DATA_BLOCK "DI_GC02_FB06_Conv_G115D"
{ S7_Optimized_Access := 'TRUE' }
VERSION : 0.1
NON_RETAIN
"FB_Conv_G115D"

BEGIN

END_DATA_BLOCK

DATA_BLOCK "DB_IO"
{ S7_Optimized_Access := 'FALSE' }
VERSION : 0.1
NON_RETAIN
   STRUCT
      CC01 : "UDT_MCC_IO";
      Power_Meter : "UDT_PAC_HW_Interface";
      UPS : "UDT_UPS_HW_Input";
      AC01 : "UDT_AC01_IO";
      AC02 : "UDT_AC02_IO";
      AC02_NT100 : "UDT_NT100_Interface";
      AC03 : "UDT_AC03_IO";
      AC03_NT100 : "UDT_NT100_Interface";
      AC04 : "UDT_AC04_IO";
      AC04_NT100 : "UDT_NT100_Interface";
      AC05 : "UDT_AC05_IO";
      AC05_NT100 : "UDT_NT100_Interface";
      GC01_SDC01 : "UDT_SDC_4Servos_IO";
      GC01_SDC02 : "UDT_SDC_4Servos_IO";
      GC02_SDC01 : "UDT_SDC_4Servos_IO";
      GC03_SDC01 : "UDT_SDC_4Servos_IO";
      GC03_SDC02 : "UDT_SDC_10Servos_IO";
      Tipper01 : "UDT_Tipper_Interface";
      ECH01 { S7_SetPoint := 'False'} : "UDT_Echelon_Interface";
      RSL01 : "UDT_RLS_Interface";
      Tipper02 : "UDT_RLS_Interface";
      ECH02 : "UDT_Echelon_Interface";
      RSL02 : "UDT_RLS_Interface";
      SG : "UDT_Merge_Singulator_Interface";
      IBST : "UDT_NBS_Interface";
      ADTA : "UDT_ADTA_Interface";
      GC01_JP03_Jam_Addon : "UDT_Jam_Addon_IO";
      GC03_FB18_Jam_Addon : "UDT_Jam_Addon_IO";
      GC01_FB10_Jam_Addon : "UDT_Jam_Addon_IO";
      GC03_JP02_Jam_Addon : "UDT_Jam_Addon_IO";
      GC01_JP02_Jam_Addon : "UDT_Jam_Addon_IO";
      GC03_JP01_Jam_Addon : "UDT_Jam_Addon_IO";
      GC01_JP01_Jam_Addon : "UDT_Jam_Addon_IO";
      GC01_FB01_Jam_Addon : "UDT_Jam_Addon_IO";
      DT01_H01 : "UDT_TL70_IO";
      DT01_H02 : "UDT_TL70_IO";
      DT02_H01 : "UDT_TL70_IO";
      DT02_H02 : "UDT_TL70_IO";
      DT03_H01 : "UDT_TL70_IO";
      DT03_H02 : "UDT_TL70_IO";
      DT04_H01 : "UDT_TL70_IO";
      GC01_FB01_XH01 : "UDT_TL70_IO";
      GC01_FB08_XH01 : "UDT_TL70_IO";
      GC01_FB16_XH01 : "UDT_TL70_IO";
      GC01_FB21_XH01 : "UDT_TL70_IO";
      GC01_FB27_XH01 : "UDT_TL70_IO";
      GC02_FB10_XH01 : "UDT_TL70_IO";
      GC03_XH01 : "UDT_TL70_IO";
      GC03_FB08_XH01 : "UDT_TL70_IO";
      GC03_XH03 : "UDT_TL70_IO";
      GC03_XH04 : "UDT_TL70_IO";
      GC04_XH01 : "UDT_TL70_IO";
      GC04_FB07_XH01 : "UDT_TL70_IO";
      GC04_FB18_XH01 : "UDT_TL70_IO";
      GC05_RC02_XH01 : "UDT_TL70_IO";
      GC06_FB08_XH01 : "UDT_TL70_IO";
      GC07_FB02_XH01 : "UDT_TL70_IO";
      GC01_FB03_B01 : "UDT_Ray26_IO";
      GC01_FB04_B01 : "UDT_Ray26_IO";
      GC01_FB05_B01 : "UDT_Ray26_IO";
      DT01_CH01_B01 : "UDT_Ray26_IO";
      DT01_RC01_B01 : "UDT_Ray26_IO";
      GC01_FB07_B01 : "UDT_Ray26_IO";
      GC01_FB08_B01 : "UDT_Ray26_IO";
      GC01_RC09_B01 : "UDT_Ray26_IO";
      GC03_RC33_B01 : "UDT_Ray26_IO";
      GC01_RC10_B01 : "UDT_Ray26_IO";
      GC01_SK11_B01 : "UDT_Ray26_IO";
      GC01_FB12_B01 : "UDT_Ray26_IO";
      GC01_FB13_B01 : "UDT_Ray26_IO";
      GC01_FB14_B01 : "UDT_Ray26_IO";
      GC01_FB28_B01 : "UDT_Ray26_IO";
      GC01_FB29_B01 : "UDT_Ray26_IO";
      GC01_FB30_B01 : "UDT_Ray26_IO";
      GC01_FB31_B01 : "UDT_Ray26_IO";
      GC02_FB03_B01 : "UDT_Ray26_IO";
      DT02_B02 : "UDT_Ray26_IO";
      GC02_FB04_B01 : "UDT_Ray26_IO";
      DT02_B01 : "UDT_Ray26_IO";
      GC02_FB06_B01 : "UDT_Ray26_IO";
      GC02_FB07_B01 : "UDT_Ray26_IO";
      GC04_FB21_B01 : "UDT_Ray26_IO";
      GC02_FB09_B01 : "UDT_Ray26_IO";
      GC02_FB10_B01 : "UDT_Ray26_IO";
      GC02_FB11_B01 : "UDT_Ray26_IO";
      GC02_FB13_B01 : "UDT_Ray26_IO";
      GC02_FB15_B01 : "UDT_Ray26_IO";
      GC02_FB16_B01 : "UDT_Ray26_IO";
      GC02_FB17_B01 : "UDT_Ray26_IO";
      GC02_FB18_B02 : "UDT_Ray26_IO";
      GC03_RC40_B01 : "UDT_Ray26_IO";
      GC03_RC02_B02 : "UDT_Ray26_IO";
      GC03_RC41_B01 : "UDT_Ray26_IO";
      GC03_RC04_B02 : "UDT_Ray26_IO";
      GC03_FB42_B01 : "UDT_Ray26_IO";
      GC03_FB09_B01 : "UDT_Ray26_IO";
      GC03_CH01_B02 : "UDT_Ray26_IO";
      DT03_B02 : "UDT_Ray26_IO";
      GC03_FB11_B01 : "UDT_Ray26_IO";
      DT03_B01 : "UDT_Ray26_IO";
      GC03_FB13_B01 : "UDT_Ray26_IO";
      GC03_FB14_B01 : "UDT_Ray26_IO";
      GC03_FB15_B01 : "UDT_Ray26_IO";
      GC03_FB16_B01 : "UDT_Ray26_IO";
      GC03_FB17_B01 : "UDT_Ray26_IO";
      GC03_FB18_B01 : "UDT_Ray26_IO";
      GC03_RC19_B01 : "UDT_Ray26_IO";
      GC03_FB21_B01 : "UDT_Ray26_IO";
      GC03_FB22_B01 : "UDT_Ray26_IO";
      GC03_FB23_B01 : "UDT_Ray26_IO";
      GC03_FB24_B01 : "UDT_Ray26_IO";
      GC03_FB25_B01 : "UDT_Ray26_IO";
      GC03_FB26_B01 : "UDT_Ray26_IO";
      GC03_FB27_B01 : "UDT_Ray26_IO";
      GC03_FB28_B01 : "UDT_Ray26_IO";
      GC03_FB29_B01 : "UDT_Ray26_IO";
      GC03_FB30_B01 : "UDT_Ray26_IO";
      GC03_FB31_B01 : "UDT_Ray26_IO";
      GC03_FB32_B01 : "UDT_Ray26_IO";
      GC03_RC33_B02 : "UDT_Ray26_IO";
      GC04_FB05_B01 : "UDT_Ray26_IO";
      GC04_FB06_B01 : "UDT_Ray26_IO";
      GC04_FB08_B01 : "UDT_Ray26_IO";
      GC04_FB09_B01 : "UDT_Ray26_IO";
      GC04_FB11_B01 : "UDT_Ray26_IO";
      GC04_FB13_B01 : "UDT_Ray26_IO";
      GC04_FB14_B01 : "UDT_Ray26_IO";
      GC04_CH01_B02 : "UDT_Ray26_IO";
      DT04_B01 : "UDT_Ray26_IO";
      GC04_FB15_B01 : "UDT_Ray26_IO";
      GC04_FB16_B01 : "UDT_Ray26_IO";
      GC04_FB17_B01 : "UDT_Ray26_IO";
      GC04_FB18_B01 : "UDT_Ray26_IO";
      GC04_FB19_B01 : "UDT_Ray26_IO";
      GC04_RC20_B01 : "UDT_Ray26_IO";
      GC05_RC02_B01 : "UDT_Ray26_IO";
      GC05_RC03_B01 : "UDT_Ray26_IO";
      GC05_FB04_B01 : "UDT_Ray26_IO";
      GC05_FB05_B01 : "UDT_Ray26_IO";
      GC05_RC06_B01 : "UDT_Ray26_IO";
      GC06_FB02_B01 : "UDT_Ray26_IO";
      GC06_FB03_B01 : "UDT_Ray26_IO";
      GC06_RC04_B01 : "UDT_Ray26_IO";
      GC06_FB05_B01 : "UDT_Ray26_IO";
      GC01_FB01_B01 : "UDT_GL2S_IO";
      GC01_FB02_B01 : "UDT_GL2S_IO";
      GC01_FB15_B01 : "UDT_GL2S_IO";
      GC01_FB16_B01 : "UDT_GL2S_IO";
      GC01_FB17_B01 : "UDT_GL2S_IO";
      GC01_FB18_B01 : "UDT_GL2S_IO";
      GC01_FB19_B01 : "UDT_GL2S_IO";
      GC01_FB20_B01 : "UDT_GL2S_IO";
      GC01_FB21_B01 : "UDT_GL2S_IO";
      GC01_FB22_B01 : "UDT_GL2S_IO";
      GC01_FB23_B01 : "UDT_GL2S_IO";
      GC01_FB24_B01 : "UDT_GL2S_IO";
      GC01_FB25_B01 : "UDT_GL2S_IO";
      GC01_FB26_B01 : "UDT_GL2S_IO";
      GC01_FB32_B01 : "UDT_GL2S_IO";
      GC02_FB01_B01 : "UDT_GL2S_IO";
      GC02_FB02_B01 : "UDT_GL2S_IO";
      GC03_CH01_B01 : "UDT_GL2S_IO";
      GC03_CH01_B03 : "UDT_GL2S_IO";
      GC03_HB05_B01 : "UDT_GL2S_IO";
      GC03_FB08_B01 : "UDT_GL2S_IO";
      GC03_FB09_B02 : "UDT_GL2S_IO";
      GC03_FB21_B02 : "UDT_GL2S_IO";
      GC03_RC33_B03 : "UDT_GL2S_IO";
      GC04_CH01_B01 : "UDT_GL2S_IO";
      GC04_CH01_B03 : "UDT_GL2S_IO";
      GC04_FB09_B02 : "UDT_GL2S_IO";
      GC06_FB05_B02 : "UDT_GL2S_IO";
      GC06_FB06_B01 : "UDT_GL2S_IO";
      GC06_FB07_B01 : "UDT_GL2S_IO";
      GC06_RC04_B02 : "UDT_GL2S_IO";
      GC06_SK08_B01 : "UDT_GL2S_IO";
      GC07_CH01_B01 : "UDT_GL2S_IO";
      GC07_CH01_B02 : "UDT_GL2S_IO";
      GC07_CH02_B01 : "UDT_GL2S_IO";
      GC07_CH02_B02 : "UDT_GL2S_IO";
      GC07_FB01_B01 : "UDT_GL2S_IO";
      GC07_FB09_B01 : "UDT_GL2S_IO";
      GC07_RC02_B02 : "UDT_GL2S_IO";
      GC07_RC03_B01 : "UDT_GL2S_IO";
      GC07_RC04_B01 : "UDT_GL2S_IO";
      GC07_RC05_B01 : "UDT_GL2S_IO";
      GC07_RC06_B01 : "UDT_GL2S_IO";
      GC07_RC07_B01 : "UDT_GL2S_IO";
      GC07_RC08_B01 : "UDT_GL2S_IO";
      GC07_RC10_B01 : "UDT_GL2S_IO";
      GC07_RC11_B01 : "UDT_GL2S_IO";
      GC01_RC06_A01 : "UDT_MultiControl_HW_Interface";
      GC01_RC09_A01 : "UDT_MultiControl_HW_Interface";
      GC01_RC10_A01 : "UDT_MultiControl_HW_Interface";
      GC02_RC05_A01 : "UDT_MultiControl_HW_Interface";
      GC03_RC01_A01 : "UDT_MultiControl_HW_Interface";
      GC03_RC02_A01 : "UDT_MultiControl_HW_Interface";
      GC03_RC03_A01 : "UDT_MultiControl_HW_Interface";
      GC03_RC04_A01 : "UDT_MultiControl_HW_Interface";
      GC03_RC20_A01 : "UDT_MultiControl_HW_Interface";
      GC03_RC20_A02 : "UDT_MultiControl_HW_Interface";
      GC04_RC20_A01 : "UDT_MultiControl_HW_Interface";
      GC05_RC01_A01 : "UDT_MultiControl_HW_Interface";
      GC05_RC02_A01 : "UDT_MultiControl_HW_Interface";
      GC05_RC02_A02 : "UDT_MultiControl_HW_Interface";
      GC05_RC02_A03 : "UDT_MultiControl_HW_Interface";
      GC05_RC03_A01 : "UDT_MultiControl_HW_Interface";
      GC05_RC06_A01 : "UDT_MultiControl_HW_Interface";
      GC06_RC01_A01 : "UDT_MultiControl_HW_Interface";
      GC07_RC03_A01 : "UDT_MultiControl_HW_Interface";
      GC07_RC04_A01 : "UDT_MultiControl_HW_Interface";
      GC07_RC04_A02 : "UDT_MultiControl_HW_Interface";
      GC07_RC05_A01 : "UDT_MultiControl_HW_Interface";
      GC07_RC06_A01 : "UDT_MultiControl_HW_Interface";
      GC07_RC07_A01 : "UDT_MultiControl_HW_Interface";
      GC07_RC07_A02 : "UDT_MultiControl_HW_Interface";
      GC07_RC07_A03 : "UDT_MultiControl_HW_Interface";
      GC07_RC08_A01 : "UDT_MultiControl_HW_Interface";
      MultiControl_Dummy : "UDT_MultiControl_HW_Interface";
      GC01_FB01 { S7_SetPoint := 'False'} : "UDT_G115D_HW_Interface";
      GC01_FB02 : "UDT_G115D_HW_Interface";
      GC01_FB03 : "UDT_G115D_HW_Interface";
      GC01_FB04 : "UDT_S210_HW_Interface";
      GC01_FB05 : "UDT_S210_HW_Interface";
      DT01 : "UDT_SWS_Interface";
      GC01_FB07 : "UDT_G115D_HW_Interface";
      GC01_FB08 : "UDT_G115D_HW_Interface";
      GC01_SK11 : "UDT_G115D_HW_Interface";
      GC01_FB12 : "UDT_S210_HW_Interface";
      GC01_FB13 : "UDT_S210_HW_Interface";
      GC01_FB14 : "UDT_S210_HW_Interface";
      GC01_FB15 : "UDT_G115D_HW_Interface";
      GC01_FB16 : "UDT_G115D_HW_Interface";
      GC01_FB17 : "UDT_G115D_HW_Interface";
      GC01_FB18 : "UDT_G115D_HW_Interface";
      GC01_FB19 : "UDT_G115D_HW_Interface";
      GC01_FB20 : "UDT_G115D_HW_Interface";
      GC01_FB21 : "UDT_G115D_HW_Interface";
      GC01_FB22 : "UDT_G115D_HW_Interface";
      GC01_FB23 : "UDT_G115D_HW_Interface";
      GC01_FB24 : "UDT_G115D_HW_Interface";
      GC01_FB25 : "UDT_G115D_HW_Interface";
      GC01_FB26 : "UDT_G115D_HW_Interface";
      GC01_FB27 : "UDT_G115D_HW_Interface";
      GC01_FB28 : "UDT_S210_HW_Interface";
      GC01_FB29 : "UDT_S210_HW_Interface";
      GC01_FB30 : "UDT_S210_HW_Interface";
      GC01_FB31 : "UDT_S210_HW_Interface";
      GC01_FB32 : "UDT_G115D_HW_Interface";
      GC02_FB01 : "UDT_G115D_HW_Interface";
      GC02_FB02 : "UDT_G115D_HW_Interface";
      GC02_FB03 : "UDT_S210_HW_Interface";
      GC02_FB04 : "UDT_S210_HW_Interface";
      DT02 : "UDT_SWS_Interface";
      GC02_FB06 : "UDT_G115D_HW_Interface";
      GC02_FB07 : "UDT_G115D_HW_Interface";
      GC02_FB08 : "UDT_G115D_HW_Interface";
      GC02_FB09 : "UDT_G115D_HW_Interface";
      GC02_FB10 : "UDT_G115D_HW_Interface";
      GC02_FB11 : "UDT_G115D_HW_Interface";
      GC02_FB12 : "UDT_G115D_HW_Interface";
      GC02_FB13 : "UDT_G115D_HW_Interface";
      GC02_FB14 : "UDT_G115D_HW_Interface";
      GC02_SK15 : "UDT_G115D_HW_Interface";
      GC02_FB16 : "UDT_S210_HW_Interface";
      GC02_FB17 : "UDT_S210_HW_Interface";
      GC02_FB18 : "UDT_S210_HW_Interface";
      GC03_HB05_M01 : "UDT_S210_HW_Interface";
      GC03_HB05_M02 : "UDT_S210_HW_Interface";
      GC03_HB05_M03 : "UDT_S210_HW_Interface";
      GC03_HB05_M04 : "UDT_S210_HW_Interface";
      GC03_HB05_M05 : "UDT_S210_HW_Interface";
      GC03_HB05_M06 : "UDT_S210_HW_Interface";
      GC03_HB05_M07 : "UDT_S210_HW_Interface";
      GC03_HB05_M08 : "UDT_S210_HW_Interface";
      GC03_HB05_M09 : "UDT_S210_HW_Interface";
      GC03_HB05_M10 : "UDT_S210_HW_Interface";
      GC03_FB06 : "UDT_G115D_HW_Interface";
      GC03_FB42 : "UDT_G115D_HW_Interface";
      GC03_FB07 : "UDT_G115D_HW_Interface";
      GC03_FB08 : "UDT_G115D_HW_Interface";
      GC03_FB09 : "UDT_G115D_HW_Interface";
      GC03_FB10 : "UDT_S210_HW_Interface";
      GC03_FB11 : "UDT_S210_HW_Interface";
      DT03 : "UDT_SWS_Interface";
      GC03_FB13 : "UDT_G115D_HW_Interface";
      GC03_FB14 : "UDT_S210_HW_Interface";
      GC03_FB15 : "UDT_S210_HW_Interface";
      GC03_FB16 : "UDT_S210_HW_Interface";
      GC03_FB17 : "UDT_S210_HW_Interface";
      GC03_FB18 : "UDT_G115D_HW_Interface";
      GC03_RC19 : "UDT_G115D_HW_Interface";
      GC03_FB21 : "UDT_G115D_HW_Interface";
      GC03_FB22 : "UDT_G115D_HW_Interface";
      GC03_FB23 : "UDT_G115D_HW_Interface";
      GC03_FB24 : "UDT_G115D_HW_Interface";
      GC03_FB25 : "UDT_G115D_HW_Interface";
      GC03_FB26 : "UDT_G115D_HW_Interface";
      GC03_FB27 : "UDT_G115D_HW_Interface";
      GC03_FB28 : "UDT_G115D_HW_Interface";
      GC03_FB29 : "UDT_G115D_HW_Interface";
      GC03_FB30 : "UDT_G115D_HW_Interface";
      GC03_FB31 : "UDT_G115D_HW_Interface";
      GC03_FB32 : "UDT_G115D_HW_Interface";
      GC03_RC33_M01 : "UDT_G115D_HW_Interface";
      GC03_RC33_M02 : "UDT_G115D_HW_Interface";
      GC04_FB04 : "UDT_G115D_HW_Interface";
      GC04_FB05 : "UDT_G115D_HW_Interface";
      GC04_FB06 : "UDT_G115D_HW_Interface";
      GC04_FB07 : "UDT_G115D_HW_Interface";
      GC04_FB08 : "UDT_G115D_HW_Interface";
      GC04_FB09 : "UDT_G115D_HW_Interface";
      GC04_FB10 : "UDT_S210_HW_Interface";
      GC04_FB11 : "UDT_S210_HW_Interface";
      DT04 : "UDT_SWS_Interface";
      GC04_FB12 : "UDT_G115D_HW_Interface";
      GC04_FB13 : "UDT_G115D_HW_Interface";
      GC04_FB14 : "UDT_G115D_HW_Interface";
      GC04_FB15 : "UDT_G115D_HW_Interface";
      GC04_FB16 : "UDT_G115D_HW_Interface";
      GC04_FB17 : "UDT_G115D_HW_Interface";
      GC04_FB18 : "UDT_G115D_HW_Interface";
      GC04_FB19 : "UDT_G115D_HW_Interface";
      GC04_RC21_M01 : "UDT_G115D_HW_Interface";
      GC04_RC21_M02 : "UDT_G115D_HW_Interface";
      GC05_FB04 : "UDT_G115D_HW_Interface";
      GC05_FB05 : "UDT_G115D_HW_Interface";
      GC05_RC07 : "UDT_G115D_HW_Interface";
      GC06_FB02 : "UDT_G115D_HW_Interface";
      GC06_FB03 : "UDT_G115D_HW_Interface";
      GC06_RC04 : "UDT_G115D_HW_Interface";
      GC06_FB05 : "UDT_G115D_HW_Interface";
      GC06_FB06 : "UDT_G115D_HW_Interface";
      GC06_FB07 : "UDT_G115D_HW_Interface";
      GC06_SK08 : "UDT_G115D_HW_Interface";
      GC07_FB01 : "UDT_G115D_HW_Interface";
      GC07_RC02_M01 : "UDT_G115D_HW_Interface";
      GC07_RC02_M02 : "UDT_G115D_HW_Interface";
      GC07_FB09 : "UDT_G115D_HW_Interface";
   END_STRUCT;


BEGIN

END_DATA_BLOCK

DATA_BLOCK "DB_System_Control"
{ S7_Optimized_Access := 'FALSE' }
VERSION : 0.1
NON_RETAIN
   STRUCT
      SSM { S7_SetPoint := 'False'} : "UDT_System_Control";
      CC01 : "UDT_System_Control";
      AC01 : "UDT_System_Control";
      AC02 : "UDT_System_Control";
      AC03 : "UDT_System_Control";
      AC04 : "UDT_System_Control";
      AC05 : "UDT_System_Control";
      GC01_SDC01 : "UDT_System_Control";
      GC01_SDC02 : "UDT_System_Control";
      GC02_SDC01 : "UDT_System_Control";
      GC03_SDC01 : "UDT_System_Control";
      GC03_SDC02 : "UDT_System_Control";
      GC03_CT01 : "UDT_System_Control";
      GC04_CT01 : "UDT_System_Control";
      Tipper01 : "UDT_System_Control";
      ECH01 : "UDT_System_Control";
      RSL01 : "UDT_System_Control";
      Tipper02 : "UDT_System_Control";
      ECH02 : "UDT_System_Control";
      RSL02 : "UDT_System_Control";
      SG : "UDT_System_Control";
      IBST : "UDT_System_Control";
      ADTA : "UDT_System_Control";
      GC01_A01 : "UDT_System_Control";
      GC01_A02 : "UDT_System_Control";
      GC01_A03 : "UDT_System_Control";
      GC01_A04 : "UDT_System_Control";
      GC01_A05 : "UDT_System_Control";
      GC02_A01 : "UDT_System_Control";
      GC02_A02 : "UDT_System_Control";
      GC02_A03 : "UDT_System_Control";
      GC03_A01 : "UDT_System_Control";
      GC03_A02 : "UDT_System_Control";
      GC03_A03 : "UDT_System_Control";
      GC03_A04 : "UDT_System_Control";
      GC03_A05 : "UDT_System_Control";
      GC03_A06 : "UDT_System_Control";
      GC04_A01 : "UDT_System_Control";
      GC04_A02 : "UDT_System_Control";
      GC04_A03 : "UDT_System_Control";
      GC05_A01 : "UDT_System_Control";
      GC06_A01 : "UDT_System_Control";
      GC07_A01 : "UDT_System_Control";
      GC01_RC06_A01 : "UDT_System_Control";
      GC01_RC09_A01 : "UDT_System_Control";
      GC01_RC10_A01 : "UDT_System_Control";
      GC02_RC05_A01 : "UDT_System_Control";
      GC03_RC01_A01 : "UDT_System_Control";
      GC03_RC02_A01 : "UDT_System_Control";
      GC03_RC03_A01 : "UDT_System_Control";
      GC03_RC04_A01 : "UDT_System_Control";
      GC03_RC20_A01 : "UDT_System_Control";
      GC03_RC20_A02 : "UDT_System_Control";
      GC04_RC20_A02 : "UDT_System_Control";
      GC05_RC01_A01 : "UDT_System_Control";
      GC05_RC02_A01 : "UDT_System_Control";
      GC05_RC02_A02 : "UDT_System_Control";
      GC05_RC02_A03 : "UDT_System_Control";
      GC05_RC03_A01 : "UDT_System_Control";
      GC05_RC06_A01 : "UDT_System_Control";
      GC06_RC01_A01 : "UDT_System_Control";
      GC07_RC03_A01 : "UDT_System_Control";
      GC07_RC04_A01 : "UDT_System_Control";
      GC07_RC04_A02 : "UDT_System_Control";
      GC07_RC05_A01 : "UDT_System_Control";
      GC07_RC06_A01 : "UDT_System_Control";
      GC07_RC07_A01 : "UDT_System_Control";
      GC07_RC07_A02 : "UDT_System_Control";
      GC07_RC07_A03 : "UDT_System_Control";
      GC07_RC08_A01 : "UDT_System_Control";
      GC01_FB01 : "UDT_System_Control";
      GC01_FB02 : "UDT_System_Control";
      GC01_FB03 : "UDT_System_Control";
      GC01_FB04 : "UDT_System_Control";
      GC01_FB05 : "UDT_System_Control";
      DT01 : "UDT_System_Control";
      GC01_RC06 : "UDT_System_Control";
      GC01_FB07 : "UDT_System_Control";
      GC01_FB08 : "UDT_System_Control";
      GC01_RC09 : "UDT_System_Control";
      GC01_RC10 : "UDT_System_Control";
      GC01_RC40 : "UDT_System_Control";
      GC01_SK11 : "UDT_System_Control";
      GC01_FB12 : "UDT_System_Control";
      GC01_FB13 : "UDT_System_Control";
      GC01_FB14 : "UDT_System_Control";
      GC01_FB15 : "UDT_System_Control";
      GC01_FB16 : "UDT_System_Control";
      GC01_FB17 : "UDT_System_Control";
      GC01_FB18 : "UDT_System_Control";
      GC01_FB19 : "UDT_System_Control";
      GC01_FB20 : "UDT_System_Control";
      GC01_FB21 : "UDT_System_Control";
      GC01_FB22 : "UDT_System_Control";
      GC01_FB23 : "UDT_System_Control";
      GC01_FB24 : "UDT_System_Control";
      GC01_FB25 : "UDT_System_Control";
      GC01_FB26 : "UDT_System_Control";
      GC01_FB27 : "UDT_System_Control";
      GC01_FB28 : "UDT_System_Control";
      GC01_FB29 : "UDT_System_Control";
      GC01_FB30 : "UDT_System_Control";
      GC01_FB31 : "UDT_System_Control";
      GC01_FB32 : "UDT_System_Control";
      GC02_FB01 : "UDT_System_Control";
      GC02_FB02 : "UDT_System_Control";
      GC02_FB03 : "UDT_System_Control";
      GC02_FB04 : "UDT_System_Control";
      DT02 : "UDT_System_Control";
      GC02_RC05 : "UDT_System_Control";
      GC02_FB06 : "UDT_System_Control";
      GC02_FB07 : "UDT_System_Control";
      GC02_FB08 : "UDT_System_Control";
      GC02_FB09 : "UDT_System_Control";
      GC02_FB10 : "UDT_System_Control";
      GC02_FB11 : "UDT_System_Control";
      GC02_FB12 : "UDT_System_Control";
      GC02_FB13 : "UDT_System_Control";
      GC02_FB14 : "UDT_System_Control";
      GC02_SK15 : "UDT_System_Control";
      GC02_FB16 : "UDT_System_Control";
      GC02_FB17 : "UDT_System_Control";
      GC02_FB18 : "UDT_System_Control";
      GC03_RC01 : "UDT_System_Control";
      GC03_RC40 : "UDT_System_Control";
      GC03_RC02 : "UDT_System_Control";
      GC03_RC03 : "UDT_System_Control";
      GC03_RC41 : "UDT_System_Control";
      GC03_RC04 : "UDT_System_Control";
      GC03_HB05 : "UDT_System_Control";
      GC03_FB06 : "UDT_System_Control";
      GC03_FB42 : "UDT_System_Control";
      GC03_FB07 : "UDT_System_Control";
      GC03_FB08 : "UDT_System_Control";
      GC03_FB09 : "UDT_System_Control";
      GC03_FB10 : "UDT_System_Control";
      GC03_FB11 : "UDT_System_Control";
      DT03 : "UDT_System_Control";
      GC03_CH01 : "UDT_System_Control";
      GC03_RC12 : "UDT_System_Control";
      GC03_FB13 : "UDT_System_Control";
      GC03_FB14 : "UDT_System_Control";
      GC03_FB15 : "UDT_System_Control";
      GC03_FB16 : "UDT_System_Control";
      GC03_FB17 : "UDT_System_Control";
      GC03_FB18 : "UDT_System_Control";
      GC03_RC19 : "UDT_System_Control";
      GC03_RC20 : "UDT_System_Control";
      GC03_FB21 : "UDT_System_Control";
      GC03_FB22 : "UDT_System_Control";
      GC03_FB23 : "UDT_System_Control";
      GC03_FB24 : "UDT_System_Control";
      GC03_FB25 : "UDT_System_Control";
      GC03_FB26 : "UDT_System_Control";
      GC03_FB27 : "UDT_System_Control";
      GC03_FB28 : "UDT_System_Control";
      GC03_FB29 : "UDT_System_Control";
      GC03_FB30 : "UDT_System_Control";
      GC03_FB31 : "UDT_System_Control";
      GC03_FB32 : "UDT_System_Control";
      GC03_RC33 : "UDT_System_Control";
      GC04_FB04 : "UDT_System_Control";
      GC04_FB05 : "UDT_System_Control";
      GC04_FB06 : "UDT_System_Control";
      GC04_FB07 : "UDT_System_Control";
      GC04_FB08 : "UDT_System_Control";
      GC04_FB09 : "UDT_System_Control";
      GC04_FB10 : "UDT_System_Control";
      GC04_FB11 : "UDT_System_Control";
      DT04 : "UDT_System_Control";
      GC04_CH01 : "UDT_System_Control";
      GC04_FB12 : "UDT_System_Control";
      GC04_FB13 : "UDT_System_Control";
      GC04_FB14 : "UDT_System_Control";
      GC04_FB15 : "UDT_System_Control";
      GC04_FB16 : "UDT_System_Control";
      GC04_FB17 : "UDT_System_Control";
      GC04_FB18 : "UDT_System_Control";
      GC04_FB19 : "UDT_System_Control";
      GC04_RC20 : "UDT_System_Control";
      GC04_RC21 : "UDT_System_Control";
      GC05_RC01 : "UDT_System_Control";
      GC05_RC02 : "UDT_System_Control";
      GC05_RC03 : "UDT_System_Control";
      GC05_RC10 : "UDT_System_Control";
      GC05_FB04 : "UDT_System_Control";
      GC05_FB05 : "UDT_System_Control";
      GC05_RC06 : "UDT_System_Control";
      GC05_RC07 : "UDT_System_Control";
      GC06_RC01 : "UDT_System_Control";
      GC06_FB02 : "UDT_System_Control";
      GC06_FB03 : "UDT_System_Control";
      GC06_RC04 : "UDT_System_Control";
      GC06_FB05 : "UDT_System_Control";
      GC06_FB06 : "UDT_System_Control";
      GC06_FB07 : "UDT_System_Control";
      GC06_SK08 : "UDT_System_Control";
      GC07_CH01 : "UDT_System_Control";
      GC07_FB01 : "UDT_System_Control";
      GC07_RC02 : "UDT_System_Control";
      GC07_RC03 : "UDT_System_Control";
      GC07_RC04 : "UDT_System_Control";
      GC07_RC05 : "UDT_System_Control";
      GC07_RC06 : "UDT_System_Control";
      GC07_RC10 : "UDT_System_Control";
      GC07_RC07 : "UDT_System_Control";
      GC07_RC08 : "UDT_System_Control";
      GC07_RC11 : "UDT_System_Control";
      GC07_CH02 : "UDT_System_Control";
      GC07_FB09 : "UDT_System_Control";
   END_STRUCT;


BEGIN

END_DATA_BLOCK

DATA_BLOCK "DI_GC02_FB03_Conv_S210"
{ S7_Optimized_Access := 'TRUE' }
VERSION : 0.1
NON_RETAIN
"FB_Conv_S210"

BEGIN

END_DATA_BLOCK

DATA_BLOCK "DB_Status"
{ S7_Optimized_Access := 'FALSE' }
AUTHOR : 'jiaqi liu'
VERSION : 0.1
NON_RETAIN
   STRUCT
      SSM : "UDT_SSM_Status";
      CC01 : "UDT_MCC_Status";
      AC01 : "UDT_AC_IO_Status";
      AC02 : "UDT_AC_SWS_Status";
      AC03 : "UDT_AC_SWS_Status";
      AC04 : "UDT_AC_SWS_Status";
      AC05 : "UDT_AC_SWS_Status";
      GC01_SDC01 : "UDT_SDC_4Servos_Status";
      GC01_SDC02 : "UDT_SDC_4Servos_Status";
      GC02_SDC01 : "UDT_SDC_4Servos_Status";
      GC03_SDC01 : "UDT_SDC_4Servos_Status";
      GC03_SDC02 : "UDT_SDC_10Servos_Status";
      GC03_CT01 : "UDT_Datalogic_AV900_Status";
      GC04_CT01 : "UDT_Datalogic_AV900_Status";
      Tipper01 : "UDT_Tipper_Status";
      ECH01 : "UDT_Echelon_Status";
      RLS01 : "UDT_RLS_Status";
      Tipper02 : "UDT_Tipper_Status";
      ECH02 : "UDT_Echelon_Status";
      RLS02 : "UDT_RLS_Status";
      SG : "UDT_Merge_Singulator_Status";
      IBST : "UDT_NBS_Status";
      ADTA : "UDT_ADTA_Status";
      GC01_A01 : "UDT_IOLink_Master_Status";
      GC01_A02 : "UDT_IOLink_Master_Status";
      GC01_A03 : "UDT_IOLink_Master_Status";
      GC01_A04 : "UDT_IOLink_Master_Status";
      GC01_A05 : "UDT_IOLink_Master_Status";
      GC02_A01 : "UDT_IOLink_Master_Status";
      GC02_A02 : "UDT_IOLink_Master_Status";
      GC02_A03 : "UDT_IOLink_Master_Status";
      GC03_A01 : "UDT_IOLink_Master_Status";
      GC03_A02 : "UDT_IOLink_Master_Status";
      GC03_A03 : "UDT_IOLink_Master_Status";
      GC03_A04 : "UDT_IOLink_Master_Status";
      GC03_A05 : "UDT_IOLink_Master_Status";
      GC03_A06 : "UDT_IOLink_Master_Status";
      GC04_A01 : "UDT_IOLink_Master_Status";
      GC04_A02 : "UDT_IOLink_Master_Status";
      GC04_A03 : "UDT_IOLink_Master_Status";
      GC05_A01 : "UDT_IOLink_Master_Status";
      GC06_A01 : "UDT_IOLink_Master_Status";
      GC07_A01 : "UDT_IOLink_Master_Status";
      GC01_RC06_A01 : "UDT_MultiControl_Status";
      GC01_RC09_A01 : "UDT_MultiControl_Status";
      GC01_RC10_A01 : "UDT_MultiControl_Status";
      GC02_RC05_A01 : "UDT_MultiControl_Status";
      GC03_RC01_A01 : "UDT_MultiControl_Status";
      GC03_RC02_A01 : "UDT_MultiControl_Status";
      GC03_RC03_A01 : "UDT_MultiControl_Status";
      GC03_RC04_A01 : "UDT_MultiControl_Status";
      GC03_RC20_A01 : "UDT_MultiControl_Status";
      GC03_RC20_A02 : "UDT_MultiControl_Status";
      GC04_RC20_A02 : "UDT_MultiControl_Status";
      GC05_RC01_A01 : "UDT_MultiControl_Status";
      GC05_RC02_A01 : "UDT_MultiControl_Status";
      GC05_RC02_A02 : "UDT_MultiControl_Status";
      GC05_RC02_A03 : "UDT_MultiControl_Status";
      GC05_RC03_A01 : "UDT_MultiControl_Status";
      GC05_RC06_A01 : "UDT_MultiControl_Status";
      GC06_RC01_A01 : "UDT_MultiControl_Status";
      GC07_RC03_A01 : "UDT_MultiControl_Status";
      GC07_RC04_A01 : "UDT_MultiControl_Status";
      GC07_RC04_A02 : "UDT_MultiControl_Status";
      GC07_RC05_A01 : "UDT_MultiControl_Status";
      GC07_RC06_A01 : "UDT_MultiControl_Status";
      GC07_RC07_A01 : "UDT_MultiControl_Status";
      GC07_RC07_A02 : "UDT_MultiControl_Status";
      GC07_RC07_A03 : "UDT_MultiControl_Status";
      GC07_RC08_A01 : "UDT_MultiControl_Status";
      GC01_FB01 : "UDT_Conv_G115D_Status";
      GC01_FB02 : "UDT_Conv_G115D_Status";
      GC01_FB03 : "UDT_Conv_G115D_Status";
      GC01_FB04 : "UDT_Conv_S210_Status";
      GC01_FB05 : "UDT_Conv_S210_Status";
      DT01 : "UDT_Conv_SWS_Status";
      GC01_RC06 : "UDT_Conv_MultiControl_Status";
      GC01_FB07 : "UDT_Conv_G115D_Status";
      GC01_FB08 : "UDT_Conv_G115D_Status";
      GC01_RC09 : "UDT_Conv_MultiControl_Status";
      GC01_RC10 : "UDT_Conv_MultiControl_Status";
      GC01_RC40 : "UDT_Conv_MultiControl_Status";
      GC01_SK11 : "UDT_Conv_G115D_Status";
      GC01_FB12 : "UDT_Conv_S210_Status";
      GC01_FB13 : "UDT_Conv_S210_Status";
      GC01_FB14 : "UDT_Conv_S210_Status";
      GC01_FB15 : "UDT_Conv_G115D_Status";
      GC01_FB16 : "UDT_Conv_G115D_Status";
      GC01_FB17 : "UDT_Conv_G115D_Status";
      GC01_FB18 : "UDT_Conv_G115D_Status";
      GC01_FB19 : "UDT_Conv_G115D_Status";
      GC01_FB20 : "UDT_Conv_G115D_Status";
      GC01_FB21 : "UDT_Conv_G115D_Status";
      GC01_FB22 : "UDT_Conv_G115D_Status";
      GC01_FB23 : "UDT_Conv_G115D_Status";
      GC01_FB24 : "UDT_Conv_G115D_Status";
      GC01_FB25 : "UDT_Conv_G115D_Status";
      GC01_FB26 : "UDT_Conv_G115D_Status";
      GC01_FB27 : "UDT_Conv_G115D_Status";
      GC01_FB28 : "UDT_Conv_S210_Status";
      GC01_FB29 : "UDT_Conv_S210_Status";
      GC01_FB30 : "UDT_Conv_S210_Status";
      GC01_FB31 : "UDT_Conv_S210_Status";
      GC01_FB32 : "UDT_Conv_G115D_Status";
      GC02_FB01 : "UDT_Conv_G115D_Status";
      GC02_FB02 : "UDT_Conv_G115D_Status";
      GC02_FB03 : "UDT_Conv_S210_Status";
      GC02_FB04 : "UDT_Conv_S210_Status";
      DT02 : "UDT_Conv_SWS_Status";
      GC02_RC05 : "UDT_Conv_MultiControl_Status";
      GC02_FB06 : "UDT_Conv_G115D_Status";
      GC02_FB07 : "UDT_Conv_G115D_Status";
      GC02_FB08 : "UDT_Conv_G115D_Status";
      GC02_FB09 : "UDT_Conv_G115D_Status";
      GC02_FB10 : "UDT_Conv_G115D_Status";
      GC02_FB11 : "UDT_Conv_G115D_Status";
      GC02_FB12 : "UDT_Conv_G115D_Status";
      GC02_FB13 : "UDT_Conv_G115D_Status";
      GC02_FB14 : "UDT_Conv_G115D_Status";
      GC02_SK15 : "UDT_Conv_G115D_Status";
      GC02_FB16 : "UDT_Conv_S210_Status";
      GC02_FB17 : "UDT_Conv_S210_Status";
      GC02_FB18 : "UDT_Conv_S210_Status";
      GC03_RC01 : "UDT_Conv_MultiControl_Status";
      GC03_RC40 : "UDT_Conv_MultiControl_Status";
      GC03_RC02 : "UDT_Conv_MultiControl_Status";
      GC03_RC03 : "UDT_Conv_MultiControl_Status";
      GC03_RC41 : "UDT_Conv_MultiControl_Status";
      GC03_RC04 : "UDT_Conv_MultiControl_Status";
      GC03_HB05 : "UDT_Conv_Multiple_S210_Status";
      GC03_FB06 : "UDT_Conv_G115D_Status";
      GC03_FB42 : "UDT_Conv_G115D_Status";
      GC03_FB07 : "UDT_Conv_G115D_Status";
      GC03_FB08 : "UDT_Conv_G115D_Status";
      GC03_FB09 : "UDT_Conv_G115D_Status";
      GC03_FB10 : "UDT_Conv_S210_Status";
      GC03_FB11 : "UDT_Conv_S210_Status";
      DT03 : "UDT_Conv_SWS_Status";
      GC03_CH01 : "UDT_Chute_Status";
      GC03_RC12 : "UDT_Conv_MultiControl_Status";
      GC03_FB13 : "UDT_Conv_G115D_Status";
      GC03_FB14 : "UDT_Conv_S210_Status";
      GC03_FB15 : "UDT_Conv_S210_Status";
      GC03_FB16 : "UDT_Conv_S210_Status";
      GC03_FB17 : "UDT_Conv_S210_Status";
      GC03_FB18 : "UDT_Conv_G115D_Status";
      GC03_RC19 : "UDT_Conv_G115D_Status";
      GC03_RC20 : "UDT_Conv_MultiControl_Status";
      GC03_FB21 : "UDT_Conv_G115D_Status";
      GC03_FB22 : "UDT_Conv_G115D_Status";
      GC03_FB23 : "UDT_Conv_G115D_Status";
      GC03_FB24 : "UDT_Conv_G115D_Status";
      GC03_FB25 : "UDT_Conv_G115D_Status";
      GC03_FB26 : "UDT_Conv_G115D_Status";
      GC03_FB27 : "UDT_Conv_G115D_Status";
      GC03_FB28 : "UDT_Conv_G115D_Status";
      GC03_FB29 : "UDT_Conv_G115D_Status";
      GC03_FB30 : "UDT_Conv_G115D_Status";
      GC03_FB31 : "UDT_Conv_G115D_Status";
      GC03_FB32 : "UDT_Conv_G115D_Status";
      GC03_RC33 : "UDT_Conv_Dual_G115D_Status";
      GC04_FB04 : "UDT_Conv_G115D_Status";
      GC04_FB05 : "UDT_Conv_G115D_Status";
      GC04_FB06 : "UDT_Conv_G115D_Status";
      GC04_FB07 : "UDT_Conv_G115D_Status";
      GC04_FB08 : "UDT_Conv_G115D_Status";
      GC04_FB09 : "UDT_Conv_G115D_Status";
      GC04_FB10 : "UDT_Conv_S210_Status";
      GC04_FB11 : "UDT_Conv_S210_Status";
      DT04 : "UDT_Conv_SWS_Status";
      GC04_CH01 { S7_SetPoint := 'False'} : "UDT_Chute_Status";
      GC04_FB12 : "UDT_Conv_G115D_Status";
      GC04_FB13 : "UDT_Conv_G115D_Status";
      GC04_FB14 : "UDT_Conv_G115D_Status";
      GC04_FB15 : "UDT_Conv_G115D_Status";
      GC04_FB16 : "UDT_Conv_G115D_Status";
      GC04_FB17 : "UDT_Conv_G115D_Status";
      GC04_FB18 : "UDT_Conv_G115D_Status";
      GC04_FB19 : "UDT_Conv_G115D_Status";
      GC04_RC20 : "UDT_Conv_MultiControl_Status";
      GC04_RC21 : "UDT_Conv_Dual_G115D_Status";
      GC05_RC01 : "UDT_Conv_MultiControl_Status";
      GC05_RC02 : "UDT_Conv_MultiControl_Status";
      GC05_RC03 : "UDT_Conv_MultiControl_Status";
      GC05_RC10 : "UDT_Conv_MultiControl_Status";
      GC05_FB04 : "UDT_Conv_G115D_Status";
      GC05_FB05 : "UDT_Conv_G115D_Status";
      GC05_RC06 : "UDT_Conv_MultiControl_Status";
      GC05_RC07 : "UDT_Conv_G115D_Status";
      GC06_RC01 : "UDT_Conv_MultiControl_Status";
      GC06_FB02 : "UDT_Conv_G115D_Status";
      GC06_FB03 : "UDT_Conv_G115D_Status";
      GC06_RC04 : "UDT_Conv_Triple_G115D_Status";
      GC06_FB05 : "UDT_Conv_G115D_Status";
      GC06_FB06 : "UDT_Conv_G115D_Status";
      GC06_FB07 : "UDT_Conv_G115D_Status";
      GC06_SK08 : "UDT_Conv_G115D_Status";
      GC07_CH01 { S7_SetPoint := 'False'} : "UDT_Chute_Status";
      GC07_FB01 : "UDT_Conv_G115D_Status";
      GC07_RC02 : "UDT_Conv_Dual_G115D_Status";
      GC07_RC03 : "UDT_Conv_MultiControl_Status";
      GC07_RC04 : "UDT_Conv_MultiControl_Status";
      GC07_RC05 : "UDT_Conv_MultiControl_Status";
      GC07_RC06 : "UDT_Conv_MultiControl_Status";
      GC07_RC10 : "UDT_Conv_MultiControl_Status";
      GC07_RC07 : "UDT_Conv_MultiControl_Status";
      GC07_RC08 : "UDT_Conv_MultiControl_Status";
      GC07_RC11 : "UDT_Conv_MultiControl_Status";
      GC07_CH02 { S7_SetPoint := 'False'} : "UDT_Chute_Status";
      GC07_FB09 : "UDT_Conv_G115D_Status";
   END_STRUCT;


BEGIN

END_DATA_BLOCK

DATA_BLOCK "DI_GC02_FB08_Conv_G115D"
{ S7_Optimized_Access := 'TRUE' }
VERSION : 0.1
NON_RETAIN
"FB_Conv_G115D"

BEGIN

END_DATA_BLOCK

DATA_BLOCK "DI_GC04_RC21_Conv_Dual_G115D"
{ S7_Optimized_Access := 'TRUE' }
VERSION : 0.1
NON_RETAIN
"FB_Conv_Dual_G115D"

BEGIN

END_DATA_BLOCK

DATA_BLOCK "DI_GC02_RC05_Conv_MultiControl"
{ S7_Optimized_Access := 'TRUE' }
VERSION : 0.1
NON_RETAIN
"FB_Conv_MultiControl"

BEGIN

END_DATA_BLOCK

DATA_BLOCK "DB_Flow_Interface"
{ S7_Optimized_Access := 'FALSE' }
VERSION : 0.1
NON_RETAIN
   STRUCT
      Dummy { S7_SetPoint := 'False'} : "UDT_Flow_Interface";
      Upstream_Dummy { S7_SetPoint := 'False'} : "UDT_Flow_Interface";
      Downstream_Dummy : "UDT_Flow_Interface";
      Tipper01 : "UDT_Flow_Interface";
      ECH01 { S7_SetPoint := 'False'} : "UDT_Flow_Interface";
      RLS01 { S7_SetPoint := 'False'} : "UDT_Flow_Interface";
      Tipper02 : "UDT_Flow_Interface";
      ECH02 { S7_SetPoint := 'False'} : "UDT_Flow_Interface";
      RLS02 { S7_SetPoint := 'False'} : "UDT_Flow_Interface";
      SG_Left { S7_SetPoint := 'False'} : "UDT_Flow_Interface";
      SG_Right : "UDT_Flow_Interface";
      IBST { S7_SetPoint := 'False'} : "UDT_Flow_Interface";
      ADTA { S7_SetPoint := 'False'} : "UDT_Flow_Interface";
      GC03_CT01 : "UDT_Flow_Interface";
      GC04_CT01 : "UDT_Flow_Interface";
      GC01_FB01 : "UDT_Flow_Interface";
      GC01_FB02 : "UDT_Flow_Interface";
      GC01_FB03 : "UDT_Flow_Interface";
      GC01_FB04 : "UDT_Flow_Interface";
      GC01_FB05 : "UDT_Flow_Interface";
      DT01 : "UDT_Flow_Interface";
      GC01_RC06 : "UDT_Flow_Interface";
      GC01_FB07 : "UDT_Flow_Interface";
      GC01_FB08 : "UDT_Flow_Interface";
      GC01_RC09 : "UDT_Flow_Interface";
      GC01_RC10 : "UDT_Flow_Interface";
      GC01_RC40 : "UDT_Flow_Interface";
      GC01_SK11 : "UDT_Flow_Interface";
      GC01_FB12 : "UDT_Flow_Interface";
      GC01_FB13 : "UDT_Flow_Interface";
      GC01_FB14 : "UDT_Flow_Interface";
      GC01_FB15 : "UDT_Flow_Interface";
      GC01_FB16 : "UDT_Flow_Interface";
      GC01_FB17 : "UDT_Flow_Interface";
      GC01_FB18 : "UDT_Flow_Interface";
      GC01_FB19 : "UDT_Flow_Interface";
      GC01_FB20 : "UDT_Flow_Interface";
      GC01_FB21 : "UDT_Flow_Interface";
      GC01_FB22 : "UDT_Flow_Interface";
      GC01_FB23 : "UDT_Flow_Interface";
      GC01_FB24 : "UDT_Flow_Interface";
      GC01_FB25 : "UDT_Flow_Interface";
      GC01_FB26 : "UDT_Flow_Interface";
      GC01_FB27 : "UDT_Flow_Interface";
      GC01_FB28 : "UDT_Flow_Interface";
      GC01_FB29 : "UDT_Flow_Interface";
      GC01_FB30 : "UDT_Flow_Interface";
      GC01_FB31 : "UDT_Flow_Interface";
      GC01_FB32 : "UDT_Flow_Interface";
      GC02_FB01 : "UDT_Flow_Interface";
      GC02_FB02 : "UDT_Flow_Interface";
      GC02_FB03 : "UDT_Flow_Interface";
      GC02_FB04 : "UDT_Flow_Interface";
      DT02 : "UDT_Flow_Interface";
      GC02_RC05 : "UDT_Flow_Interface";
      GC02_FB06 : "UDT_Flow_Interface";
      GC02_FB07 : "UDT_Flow_Interface";
      GC02_FB08 : "UDT_Flow_Interface";
      GC02_FB09 : "UDT_Flow_Interface";
      GC02_FB10 : "UDT_Flow_Interface";
      GC02_FB11 : "UDT_Flow_Interface";
      GC02_FB12 : "UDT_Flow_Interface";
      GC02_FB13 : "UDT_Flow_Interface";
      GC02_FB14 : "UDT_Flow_Interface";
      GC02_SK15 : "UDT_Flow_Interface";
      GC02_FB16 : "UDT_Flow_Interface";
      GC02_FB17 : "UDT_Flow_Interface";
      GC02_FB18 : "UDT_Flow_Interface";
      GC03_RC01 : "UDT_Flow_Interface";
      GC03_RC40 : "UDT_Flow_Interface";
      GC03_RC02 : "UDT_Flow_Interface";
      GC03_RC02_END : "UDT_Flow_Interface";
      GC03_RC03 : "UDT_Flow_Interface";
      GC03_RC41 : "UDT_Flow_Interface";
      GC03_RC04 : "UDT_Flow_Interface";
      GC03_RC04_END : "UDT_Flow_Interface";
      GC03_HB05_Infeed : "UDT_Flow_Interface";
      GC03_HB05 : "UDT_Flow_Interface";
      GC03_FB06 : "UDT_Flow_Interface";
      GC03_FB42 : "UDT_Flow_Interface";
      GC03_FB07 : "UDT_Flow_Interface";
      GC03_FB08 : "UDT_Flow_Interface";
      GC03_FB09 : "UDT_Flow_Interface";
      GC03_FB10 : "UDT_Flow_Interface";
      GC03_FB11 : "UDT_Flow_Interface";
      DT03 : "UDT_Flow_Interface";
      GC03_CH01 : "UDT_Flow_Interface";
      GC03_RC12 : "UDT_Flow_Interface";
      GC03_FB13 : "UDT_Flow_Interface";
      GC03_FB14 : "UDT_Flow_Interface";
      GC03_FB15 : "UDT_Flow_Interface";
      GC03_FB16 : "UDT_Flow_Interface";
      GC03_FB17 : "UDT_Flow_Interface";
      GC03_FB18 : "UDT_Flow_Interface";
      GC03_FB18_END : "UDT_Flow_Interface";
      GC03_RC19 : "UDT_Flow_Interface";
      GC03_RC20 : "UDT_Flow_Interface";
      GC03_FB21 : "UDT_Flow_Interface";
      GC03_FB22 : "UDT_Flow_Interface";
      GC03_FB23 : "UDT_Flow_Interface";
      GC03_FB24 : "UDT_Flow_Interface";
      GC03_FB25 : "UDT_Flow_Interface";
      GC03_FB26 : "UDT_Flow_Interface";
      GC03_FB27 : "UDT_Flow_Interface";
      GC03_FB28 : "UDT_Flow_Interface";
      GC03_FB29 : "UDT_Flow_Interface";
      GC03_FB30 : "UDT_Flow_Interface";
      GC03_FB31 : "UDT_Flow_Interface";
      GC03_FB32 : "UDT_Flow_Interface";
      GC03_FB32_Infeed : "UDT_Flow_Interface";
      GC03_RC33 : "UDT_Flow_Interface";
      GC04_FB04 : "UDT_Flow_Interface";
      GC04_FB05 : "UDT_Flow_Interface";
      GC04_FB06 : "UDT_Flow_Interface";
      GC04_FB07 : "UDT_Flow_Interface";
      GC04_FB08 : "UDT_Flow_Interface";
      GC04_FB09 : "UDT_Flow_Interface";
      GC04_FB10 : "UDT_Flow_Interface";
      GC04_FB11 : "UDT_Flow_Interface";
      DT04 : "UDT_Flow_Interface";
      GC04_CH01 : "UDT_Flow_Interface";
      GC04_FB12 : "UDT_Flow_Interface";
      GC04_FB13 : "UDT_Flow_Interface";
      GC04_FB14 : "UDT_Flow_Interface";
      GC04_FB15 : "UDT_Flow_Interface";
      GC04_FB16 : "UDT_Flow_Interface";
      GC04_FB17 : "UDT_Flow_Interface";
      GC04_FB18 : "UDT_Flow_Interface";
      GC04_FB19 : "UDT_Flow_Interface";
      GC04_RC20 : "UDT_Flow_Interface";
      GC04_RC21 : "UDT_Flow_Interface";
      GC05_RC01 : "UDT_Flow_Interface";
      GC05_RC02 : "UDT_Flow_Interface";
      GC05_RC03 : "UDT_Flow_Interface";
      GC05_RC10 : "UDT_Flow_Interface";
      GC05_FB04 : "UDT_Flow_Interface";
      GC05_FB05 : "UDT_Flow_Interface";
      GC05_RC06 : "UDT_Flow_Interface";
      GC05_RC06_END : "UDT_Flow_Interface";
      GC05_RC07 : "UDT_Flow_Interface";
      GC06_RC01 : "UDT_Flow_Interface";
      GC06_FB02 : "UDT_Flow_Interface";
      GC06_FB03 : "UDT_Flow_Interface";
      GC06_FB03_END : "UDT_Flow_Interface";
      GC06_RC04_Infeed : "UDT_Flow_Interface";
      GC06_RC04 : "UDT_Flow_Interface";
      GC06_FB05 : "UDT_Flow_Interface";
      GC06_FB06 : "UDT_Flow_Interface";
      GC06_FB07 : "UDT_Flow_Interface";
      GC06_SK08 : "UDT_Flow_Interface";
      GC07_CH01 : "UDT_Flow_Interface";
      GC07_FB01 : "UDT_Flow_Interface";
      GC07_RC02 : "UDT_Flow_Interface";
      GC07_RC03 : "UDT_Flow_Interface";
      GC07_RC04 : "UDT_Flow_Interface";
      GC07_RC05 : "UDT_Flow_Interface";
      GC07_RC06 : "UDT_Flow_Interface";
      GC07_RC10 : "UDT_Flow_Interface";
      GC07_RC07 : "UDT_Flow_Interface";
      GC07_RC08 : "UDT_Flow_Interface";
      GC07_RC11 : "UDT_Flow_Interface";
      GC07_CH02 : "UDT_Flow_Interface";
      GC07_FB09 : "UDT_Flow_Interface";
   END_STRUCT;


BEGIN
   Upstream_Dummy.Operational := TRUE;
   Upstream_Dummy.Available := TRUE;
   Upstream_Dummy.Cascade_Startup := TRUE;
   Upstream_Dummy.Cascade_Shutdown := TRUE;
   Upstream_Dummy.Motor_Run := TRUE;
   Downstream_Dummy.RTR := TRUE;
   Downstream_Dummy.Operational := TRUE;
   Downstream_Dummy.Available := TRUE;
   Downstream_Dummy.Cascade_Startup := TRUE;
   Downstream_Dummy.Motor_Run := TRUE;
   Downstream_Dummy.Displacement := 10;

END_DATA_BLOCK

DATA_BLOCK "DI_GC02_FB09_Conv_G115D"
{ S7_Optimized_Access := 'TRUE' }
VERSION : 0.1
NON_RETAIN
"FB_Conv_G115D"

BEGIN

END_DATA_BLOCK

DATA_BLOCK "DI_GC02_FB10_Conv_G115D"
{ S7_Optimized_Access := 'TRUE' }
VERSION : 0.1
NON_RETAIN
"FB_Conv_G115D"

BEGIN

END_DATA_BLOCK

DATA_BLOCK "DI_GC02_FB11_Conv_G115D"
{ S7_Optimized_Access := 'TRUE' }
VERSION : 0.1
NON_RETAIN
"FB_Conv_G115D"

BEGIN

END_DATA_BLOCK

DATA_BLOCK "DI_GC02_FB12_Conv_G115D"
{ S7_Optimized_Access := 'TRUE' }
VERSION : 0.1
NON_RETAIN
"FB_Conv_G115D"

BEGIN

END_DATA_BLOCK

DATA_BLOCK "DI_GC02_FB13_Conv_G115D"
{ S7_Optimized_Access := 'TRUE' }
VERSION : 0.1
NON_RETAIN
"FB_Conv_G115D"

BEGIN

END_DATA_BLOCK

DATA_BLOCK "DI_GC02_FB14_Conv_G115D"
{ S7_Optimized_Access := 'TRUE' }
VERSION : 0.1
NON_RETAIN
"FB_Conv_G115D"

BEGIN

END_DATA_BLOCK

DATA_BLOCK "DB_General_Status"
{ S7_Optimized_Access := 'FALSE' }
VERSION : 0.1
NON_RETAIN
   STRUCT
      SSM : "UDT_General_Status";
      CC01 : "UDT_General_Status";
      AC01 : "UDT_General_Status";
      AC02 : "UDT_General_Status";
      AC03 : "UDT_General_Status";
      AC04 : "UDT_General_Status";
      AC05 : "UDT_General_Status";
      GC01_SDC01 : "UDT_General_Status";
      GC01_SDC02 : "UDT_General_Status";
      GC02_SDC01 : "UDT_General_Status";
      GC03_SDC01 : "UDT_General_Status";
      GC03_SDC02 : "UDT_General_Status";
      GC03_CT01 : "UDT_General_Status";
      GC04_CT01 : "UDT_General_Status";
      Tipper01 : "UDT_General_Status";
      ECH01 : "UDT_General_Status";
      RSL01 : "UDT_General_Status";
      Tipper02 : "UDT_General_Status";
      ECH02 : "UDT_General_Status";
      RSL02 : "UDT_General_Status";
      SG : "UDT_General_Status";
      IBST : "UDT_General_Status";
      ADTA : "UDT_General_Status";
      GC01_A01 : "UDT_General_Status";
      GC01_A02 : "UDT_General_Status";
      GC01_A03 : "UDT_General_Status";
      GC01_A04 : "UDT_General_Status";
      GC01_A05 : "UDT_General_Status";
      GC02_A01 : "UDT_General_Status";
      GC02_A02 : "UDT_General_Status";
      GC02_A03 : "UDT_General_Status";
      GC03_A01 : "UDT_General_Status";
      GC03_A02 : "UDT_General_Status";
      GC03_A03 : "UDT_General_Status";
      GC03_A04 : "UDT_General_Status";
      GC03_A05 : "UDT_General_Status";
      GC03_A06 : "UDT_General_Status";
      GC04_A01 : "UDT_General_Status";
      GC04_A02 : "UDT_General_Status";
      GC04_A03 : "UDT_General_Status";
      GC05_A01 : "UDT_General_Status";
      GC06_A01 : "UDT_General_Status";
      GC07_A01 : "UDT_General_Status";
      GC01_RC06_A01 : "UDT_General_Status";
      GC01_RC09_A01 : "UDT_General_Status";
      GC01_RC10_A01 : "UDT_General_Status";
      GC02_RC05_A01 : "UDT_General_Status";
      GC03_RC01_A01 : "UDT_General_Status";
      GC03_RC02_A01 : "UDT_General_Status";
      GC03_RC03_A01 : "UDT_General_Status";
      GC03_RC04_A01 : "UDT_General_Status";
      GC03_RC20_A01 : "UDT_General_Status";
      GC03_RC20_A02 : "UDT_General_Status";
      GC04_RC20_A02 : "UDT_General_Status";
      GC05_RC01_A01 : "UDT_General_Status";
      GC05_RC02_A01 : "UDT_General_Status";
      GC05_RC02_A02 : "UDT_General_Status";
      GC05_RC02_A03 : "UDT_General_Status";
      GC05_RC03_A01 : "UDT_General_Status";
      GC05_RC06_A01 : "UDT_General_Status";
      GC06_RC01_A01 : "UDT_General_Status";
      GC07_RC03_A01 : "UDT_General_Status";
      GC07_RC04_A01 : "UDT_General_Status";
      GC07_RC04_A02 : "UDT_General_Status";
      GC07_RC05_A01 : "UDT_General_Status";
      GC07_RC06_A01 : "UDT_General_Status";
      GC07_RC07_A01 : "UDT_General_Status";
      GC07_RC07_A02 : "UDT_General_Status";
      GC07_RC07_A03 : "UDT_General_Status";
      GC07_RC08_A01 : "UDT_General_Status";
      GC01_FB01 : "UDT_General_Status";
      GC01_FB02 : "UDT_General_Status";
      GC01_FB03 : "UDT_General_Status";
      GC01_FB04 : "UDT_General_Status";
      GC01_FB05 : "UDT_General_Status";
      DT01 : "UDT_General_Status";
      GC01_RC06 : "UDT_General_Status";
      GC01_FB07 : "UDT_General_Status";
      GC01_FB08 : "UDT_General_Status";
      GC01_RC09 : "UDT_General_Status";
      GC01_RC10 : "UDT_General_Status";
      GC01_RC40 : "UDT_General_Status";
      GC01_SK11 : "UDT_General_Status";
      GC01_FB12 : "UDT_General_Status";
      GC01_FB13 : "UDT_General_Status";
      GC01_FB14 : "UDT_General_Status";
      GC01_FB15 : "UDT_General_Status";
      GC01_FB16 : "UDT_General_Status";
      GC01_FB17 : "UDT_General_Status";
      GC01_FB18 : "UDT_General_Status";
      GC01_FB19 : "UDT_General_Status";
      GC01_FB20 : "UDT_General_Status";
      GC01_FB21 : "UDT_General_Status";
      GC01_FB22 : "UDT_General_Status";
      GC01_FB23 : "UDT_General_Status";
      GC01_FB24 : "UDT_General_Status";
      GC01_FB25 : "UDT_General_Status";
      GC01_FB26 : "UDT_General_Status";
      GC01_FB27 : "UDT_General_Status";
      GC01_FB28 : "UDT_General_Status";
      GC01_FB29 : "UDT_General_Status";
      GC01_FB30 : "UDT_General_Status";
      GC01_FB31 : "UDT_General_Status";
      GC01_FB32 : "UDT_General_Status";
      GC02_FB01 : "UDT_General_Status";
      GC02_FB02 : "UDT_General_Status";
      GC02_FB03 : "UDT_General_Status";
      GC02_FB04 : "UDT_General_Status";
      DT02 : "UDT_General_Status";
      GC02_RC05 : "UDT_General_Status";
      GC02_FB06 : "UDT_General_Status";
      GC02_FB07 : "UDT_General_Status";
      GC02_FB08 : "UDT_General_Status";
      GC02_FB09 : "UDT_General_Status";
      GC02_FB10 : "UDT_General_Status";
      GC02_FB11 : "UDT_General_Status";
      GC02_FB12 : "UDT_General_Status";
      GC02_FB13 : "UDT_General_Status";
      GC02_FB14 : "UDT_General_Status";
      GC02_SK15 : "UDT_General_Status";
      GC02_FB16 : "UDT_General_Status";
      GC02_FB17 : "UDT_General_Status";
      GC02_FB18 : "UDT_General_Status";
      GC03_RC01 : "UDT_General_Status";
      GC03_RC40 : "UDT_General_Status";
      GC03_RC02 : "UDT_General_Status";
      GC03_RC03 : "UDT_General_Status";
      GC03_RC41 : "UDT_General_Status";
      GC03_RC04 : "UDT_General_Status";
      GC03_HB05 : "UDT_General_Status";
      GC03_FB06 : "UDT_General_Status";
      GC03_FB42 : "UDT_General_Status";
      GC03_FB07 : "UDT_General_Status";
      GC03_FB08 : "UDT_General_Status";
      GC03_FB09 : "UDT_General_Status";
      GC03_FB10 : "UDT_General_Status";
      GC03_FB11 : "UDT_General_Status";
      DT03 : "UDT_General_Status";
      GC03_CH01 : "UDT_General_Status";
      GC03_RC12 : "UDT_General_Status";
      GC03_FB13 : "UDT_General_Status";
      GC03_FB14 : "UDT_General_Status";
      GC03_FB15 : "UDT_General_Status";
      GC03_FB16 : "UDT_General_Status";
      GC03_FB17 : "UDT_General_Status";
      GC03_FB18 : "UDT_General_Status";
      GC03_RC19 : "UDT_General_Status";
      GC03_RC20 : "UDT_General_Status";
      GC03_FB21 : "UDT_General_Status";
      GC03_FB22 : "UDT_General_Status";
      GC03_FB23 : "UDT_General_Status";
      GC03_FB24 : "UDT_General_Status";
      GC03_FB25 : "UDT_General_Status";
      GC03_FB26 : "UDT_General_Status";
      GC03_FB27 : "UDT_General_Status";
      GC03_FB28 : "UDT_General_Status";
      GC03_FB29 : "UDT_General_Status";
      GC03_FB30 : "UDT_General_Status";
      GC03_FB31 : "UDT_General_Status";
      GC03_FB32 : "UDT_General_Status";
      GC03_RC33 : "UDT_General_Status";
      GC04_FB04 : "UDT_General_Status";
      GC04_FB05 : "UDT_General_Status";
      GC04_FB06 : "UDT_General_Status";
      GC04_FB07 : "UDT_General_Status";
      GC04_FB08 : "UDT_General_Status";
      GC04_FB09 : "UDT_General_Status";
      GC04_FB10 : "UDT_General_Status";
      GC04_FB11 : "UDT_General_Status";
      DT04 : "UDT_General_Status";
      GC04_CH01 : "UDT_General_Status";
      GC04_FB12 : "UDT_General_Status";
      GC04_FB13 : "UDT_General_Status";
      GC04_FB14 : "UDT_General_Status";
      GC04_FB15 : "UDT_General_Status";
      GC04_FB16 : "UDT_General_Status";
      GC04_FB17 : "UDT_General_Status";
      GC04_FB18 : "UDT_General_Status";
      GC04_FB19 : "UDT_General_Status";
      GC04_RC20 : "UDT_General_Status";
      GC04_RC21 : "UDT_General_Status";
      GC05_RC01 : "UDT_General_Status";
      GC05_RC02 : "UDT_General_Status";
      GC05_RC03 : "UDT_General_Status";
      GC05_RC10 : "UDT_General_Status";
      GC05_FB04 : "UDT_General_Status";
      GC05_FB05 : "UDT_General_Status";
      GC05_RC06 : "UDT_General_Status";
      GC05_RC07 : "UDT_General_Status";
      GC06_RC01 : "UDT_General_Status";
      GC06_FB02 : "UDT_General_Status";
      GC06_FB03 : "UDT_General_Status";
      GC06_RC04 : "UDT_General_Status";
      GC06_FB05 : "UDT_General_Status";
      GC06_FB06 : "UDT_General_Status";
      GC06_FB07 : "UDT_General_Status";
      GC06_SK08 : "UDT_General_Status";
      GC07_CH01 : "UDT_General_Status";
      GC07_FB01 : "UDT_General_Status";
      GC07_RC02 : "UDT_General_Status";
      GC07_RC03 : "UDT_General_Status";
      GC07_RC04 : "UDT_General_Status";
      GC07_RC05 : "UDT_General_Status";
      GC07_RC06 : "UDT_General_Status";
      GC07_RC10 : "UDT_General_Status";
      GC07_RC07 : "UDT_General_Status";
      GC07_RC08 : "UDT_General_Status";
      GC07_RC11 : "UDT_General_Status";
      GC07_CH02 : "UDT_General_Status";
      GC07_FB09 : "UDT_General_Status";
   END_STRUCT;


BEGIN

END_DATA_BLOCK

DATA_BLOCK "DI_GC02_SK15_Conv_G115D"
{ S7_Optimized_Access := 'TRUE' }
VERSION : 0.1
NON_RETAIN
"FB_Conv_G115D"

BEGIN

END_DATA_BLOCK

DATA_BLOCK "DI_GC02_FB17_Conv_S210"
{ S7_Optimized_Access := 'TRUE' }
VERSION : 0.1
NON_RETAIN
"FB_Conv_S210"

BEGIN

END_DATA_BLOCK

DATA_BLOCK "DI_GC02_FB18_Conv_S210"
{ S7_Optimized_Access := 'TRUE' }
VERSION : 0.1
NON_RETAIN
"FB_Conv_S210"

BEGIN

END_DATA_BLOCK

DATA_BLOCK "DI_DT02_Conv_SWS"
{ S7_Optimized_Access := 'TRUE' }
VERSION : 0.1
NON_RETAIN
"FB_Conv_SWS"

BEGIN

END_DATA_BLOCK

DATA_BLOCK "DI_GC02_FB04_Conv_S210"
{ S7_Optimized_Access := 'TRUE' }
VERSION : 0.1
NON_RETAIN
"FB_Conv_S210"

BEGIN

END_DATA_BLOCK

DATA_BLOCK "DI_GC02_FB07_Conv_G115D"
{ S7_Optimized_Access := 'TRUE' }
VERSION : 0.1
NON_RETAIN
"FB_Conv_G115D"

BEGIN

END_DATA_BLOCK

DATA_BLOCK "DI_GC02_FB02_Conv_G115D"
{ S7_Optimized_Access := 'TRUE' }
VERSION : 0.1
NON_RETAIN
"FB_Conv_G115D"

BEGIN

END_DATA_BLOCK

DATA_BLOCK "DB_Global"
{ S7_Optimized_Access := 'TRUE' }
VERSION : 0.1
NON_RETAIN
"UDT_Global"

BEGIN

END_DATA_BLOCK

DATA_BLOCK "DI_GC02_FB01_Conv_G115D"
{ S7_Optimized_Access := 'TRUE' }
VERSION : 0.1
NON_RETAIN
"FB_Conv_G115D"

BEGIN

END_DATA_BLOCK

DATA_BLOCK "DB_External"
{ S7_Optimized_Access := 'TRUE' }
VERSION : 0.1
NON_RETAIN
   VAR
      ECH01 { S7_SetPoint := 'False'} : "UDT_External_Request";
      RLS01 { S7_SetPoint := 'False'} : "UDT_External_Request";
      ECH02 { S7_SetPoint := 'False'} : "UDT_External_Request";
      RLS02 { S7_SetPoint := 'False'} : "UDT_External_Request";
      SG01 { S7_SetPoint := 'False'} : "UDT_External_Request";
      IBST01 { S7_SetPoint := 'False'} : "UDT_External_Request";
      ADTA01 { S7_SetPoint := 'False'} : "UDT_External_Request";
      GC03_CT01 : "UDT_External_Request";
      GC04_CT01 : "UDT_External_Request";
      GC01_FB01 : "UDT_External_Request";
      GC01_FB02 : "UDT_External_Request";
      GC01_FB03 : "UDT_External_Request";
      GC01_FB04 : "UDT_External_Request";
      GC01_FB05 : "UDT_External_Request";
      DT01 : "UDT_External_Request";
      GC01_RC06 : "UDT_External_Request";
      GC01_FB07 : "UDT_External_Request";
      GC01_FB08 : "UDT_External_Request";
      GC01_RC09 : "UDT_External_Request";
      GC01_RC10 : "UDT_External_Request";
      GC01_RC40 : "UDT_External_Request";
      GC01_SK11 : "UDT_External_Request";
      GC01_FB12 : "UDT_External_Request";
      GC01_FB13 : "UDT_External_Request";
      GC01_FB14 : "UDT_External_Request";
      GC01_FB15 : "UDT_External_Request";
      GC01_FB16 : "UDT_External_Request";
      GC01_FB17 : "UDT_External_Request";
      GC01_FB18 : "UDT_External_Request";
      GC01_FB19 : "UDT_External_Request";
      GC01_FB20 : "UDT_External_Request";
      GC01_FB21 : "UDT_External_Request";
      GC01_FB22 : "UDT_External_Request";
      GC01_FB23 : "UDT_External_Request";
      GC01_FB24 : "UDT_External_Request";
      GC01_FB25 : "UDT_External_Request";
      GC01_FB26 : "UDT_External_Request";
      GC01_FB27 : "UDT_External_Request";
      GC01_FB28 : "UDT_External_Request";
      GC01_FB29 : "UDT_External_Request";
      GC01_FB30 : "UDT_External_Request";
      GC01_FB31 : "UDT_External_Request";
      GC01_FB32 : "UDT_External_Request";
      GC02_FB01 : "UDT_External_Request";
      GC02_FB02 : "UDT_External_Request";
      GC02_FB03 : "UDT_External_Request";
      GC02_FB04 : "UDT_External_Request";
      DT02 : "UDT_External_Request";
      GC02_RC05 : "UDT_External_Request";
      GC02_FB06 : "UDT_External_Request";
      GC02_FB07 : "UDT_External_Request";
      GC02_FB08 : "UDT_External_Request";
      GC02_FB09 : "UDT_External_Request";
      GC02_FB10 : "UDT_External_Request";
      GC02_FB11 : "UDT_External_Request";
      GC02_FB12 : "UDT_External_Request";
      GC02_FB13 : "UDT_External_Request";
      GC02_FB14 : "UDT_External_Request";
      GC02_SK15 : "UDT_External_Request";
      GC02_FB16 : "UDT_External_Request";
      GC02_FB17 : "UDT_External_Request";
      GC02_FB18 : "UDT_External_Request";
      GC03_RC01 : "UDT_External_Request";
      GC03_RC40 : "UDT_External_Request";
      GC03_RC02 : "UDT_External_Request";
      GC03_RC03 : "UDT_External_Request";
      GC03_RC41 : "UDT_External_Request";
      GC03_RC04 : "UDT_External_Request";
      GC03_HB05 : "UDT_External_Request";
      GC03_FB06 : "UDT_External_Request";
      GC03_FB42 : "UDT_External_Request";
      GC03_FB07 : "UDT_External_Request";
      GC03_FB08 : "UDT_External_Request";
      GC03_FB09 : "UDT_External_Request";
      GC03_FB10 : "UDT_External_Request";
      GC03_FB11 : "UDT_External_Request";
      DT03 : "UDT_External_Request";
      GC03_CH01 : "UDT_External_Request";
      GC03_RC12 : "UDT_External_Request";
      GC03_FB13 : "UDT_External_Request";
      GC03_FB14 : "UDT_External_Request";
      GC03_FB15 : "UDT_External_Request";
      GC03_FB16 : "UDT_External_Request";
      GC03_FB17 : "UDT_External_Request";
      GC03_FB18 : "UDT_External_Request";
      GC03_RC19 : "UDT_External_Request";
      GC03_RC20 : "UDT_External_Request";
      GC03_FB21 : "UDT_External_Request";
      GC03_FB22 : "UDT_External_Request";
      GC03_FB23 : "UDT_External_Request";
      GC03_FB24 : "UDT_External_Request";
      GC03_FB25 : "UDT_External_Request";
      GC03_FB26 : "UDT_External_Request";
      GC03_FB27 : "UDT_External_Request";
      GC03_FB28 : "UDT_External_Request";
      GC03_FB29 : "UDT_External_Request";
      GC03_FB30 : "UDT_External_Request";
      GC03_FB31 : "UDT_External_Request";
      GC03_FB32 : "UDT_External_Request";
      GC03_RC33 : "UDT_External_Request";
      GC04_FB04 : "UDT_External_Request";
      GC04_FB05 : "UDT_External_Request";
      GC04_FB06 : "UDT_External_Request";
      GC04_FB07 : "UDT_External_Request";
      GC04_FB08 : "UDT_External_Request";
      GC04_FB09 : "UDT_External_Request";
      GC04_FB10 : "UDT_External_Request";
      GC04_FB11 : "UDT_External_Request";
      DT04 : "UDT_External_Request";
      GC04_CH01 : "UDT_External_Request";
      GC04_FB12 : "UDT_External_Request";
      GC04_FB13 : "UDT_External_Request";
      GC04_FB14 : "UDT_External_Request";
      GC04_FB15 : "UDT_External_Request";
      GC04_FB16 : "UDT_External_Request";
      GC04_FB17 : "UDT_External_Request";
      GC04_FB18 : "UDT_External_Request";
      GC04_FB19 : "UDT_External_Request";
      GC04_RC20 : "UDT_External_Request";
      GC04_RC21 : "UDT_External_Request";
      GC05_RC01 : "UDT_External_Request";
      GC05_RC02 : "UDT_External_Request";
      GC05_RC03 : "UDT_External_Request";
      GC05_RC10 : "UDT_External_Request";
      GC05_FB04 : "UDT_External_Request";
      GC05_FB05 : "UDT_External_Request";
      GC05_RC06 : "UDT_External_Request";
      GC05_RC07 : "UDT_External_Request";
      GC06_RC01 : "UDT_External_Request";
      GC06_FB02 : "UDT_External_Request";
      GC06_FB03 : "UDT_External_Request";
      GC06_RC04 : "UDT_External_Request";
      GC06_FB05 : "UDT_External_Request";
      GC06_FB06 : "UDT_External_Request";
      GC06_FB07 : "UDT_External_Request";
      GC06_SK08 : "UDT_External_Request";
      GC07_CH01 : "UDT_External_Request";
      GC07_FB01 : "UDT_External_Request";
      GC07_RC02 : "UDT_External_Request";
      GC07_RC03 : "UDT_External_Request";
      GC07_RC04 : "UDT_External_Request";
      GC07_RC05 : "UDT_External_Request";
      GC07_RC06 : "UDT_External_Request";
      GC07_RC10 : "UDT_External_Request";
      GC07_RC07 : "UDT_External_Request";
      GC07_RC08 : "UDT_External_Request";
      GC07_RC11 : "UDT_External_Request";
      GC07_CH02 : "UDT_External_Request";
      GC07_FB09 : "UDT_External_Request";
   END_VAR


BEGIN

END_DATA_BLOCK

DATA_BLOCK "DB_Command"
{ S7_Optimized_Access := 'FALSE' }
AUTHOR : 'jiaqi liu'
VERSION : 0.1
   STRUCT
      CC01 { S7_SetPoint := 'False'} : "UDT_MCC_Command";
      SCADA { S7_SetPoint := 'False'} : "UDT_SCADA_Command";
      HMI { S7_SetPoint := 'False'} : "UDT_HMI_Command";
      Tipper01 { S7_SetPoint := 'False'} : "UDT_Tipper_Command";
      ECH01 { S7_SetPoint := 'False'} : "UDT_Echelon_Command";
      RLS01 { S7_SetPoint := 'False'} : "UDT_RLS_Command";
      Tipper02 : "UDT_Tipper_Command";
      ECH02 { S7_SetPoint := 'False'} : "UDT_Echelon_Command";
      RLS02 { S7_SetPoint := 'False'} : "UDT_RLS_Command";
      SG { S7_SetPoint := 'False'} : "UDT_Merge_Singulator_Command";
      IBST { S7_SetPoint := 'False'} : "UDT_NBS_Command";
      ADTA { S7_SetPoint := 'False'} : "UDT_ADTA_Command";
      GC03_CT01 { S7_SetPoint := 'False'} : "UDT_Datalogic_AV900_Command";
      GC04_CT01 : "UDT_Datalogic_AV900_Command";
      GC01_A01 { S7_SetPoint := 'False'} : "UDT_IOLink_Master_Command";
      GC01_A02 : "UDT_IOLink_Master_Command";
      GC01_A03 : "UDT_IOLink_Master_Command";
      GC01_A04 : "UDT_IOLink_Master_Command";
      GC01_A05 : "UDT_IOLink_Master_Command";
      GC02_A01 : "UDT_IOLink_Master_Command";
      GC02_A02 : "UDT_IOLink_Master_Command";
      GC02_A03 : "UDT_IOLink_Master_Command";
      GC03_A01 : "UDT_IOLink_Master_Command";
      GC03_A02 : "UDT_IOLink_Master_Command";
      GC03_A03 : "UDT_IOLink_Master_Command";
      GC03_A04 : "UDT_IOLink_Master_Command";
      GC03_A05 : "UDT_IOLink_Master_Command";
      GC03_A06 : "UDT_IOLink_Master_Command";
      GC04_A01 : "UDT_IOLink_Master_Command";
      GC04_A02 : "UDT_IOLink_Master_Command";
      GC04_A03 : "UDT_IOLink_Master_Command";
      GC05_A01 : "UDT_IOLink_Master_Command";
      GC06_A01 : "UDT_IOLink_Master_Command";
      GC07_A01 : "UDT_IOLink_Master_Command";
      GC01_FB01 { S7_SetPoint := 'False'} : "UDT_Conv_G115D_Command";
      GC01_FB02 : "UDT_Conv_G115D_Command";
      GC01_FB03 : "UDT_Conv_G115D_Command";
      GC01_FB04 : "UDT_Conv_S210_Command";
      GC01_FB05 : "UDT_Conv_S210_Command";
      DT01 : "UDT_Conv_SWS_Command";
      GC01_RC06 : "UDT_Conv_MultiControl_Command";
      GC01_FB07 : "UDT_Conv_G115D_Command";
      GC01_FB08 : "UDT_Conv_G115D_Command";
      GC01_RC09 : "UDT_Conv_MultiControl_Command";
      GC01_RC10 : "UDT_Conv_MultiControl_Command";
      GC01_RC40 : "UDT_Conv_MultiControl_Command";
      GC01_SK11 : "UDT_Conv_G115D_Command";
      GC01_FB12 : "UDT_Conv_S210_Command";
      GC01_FB13 : "UDT_Conv_S210_Command";
      GC01_FB14 : "UDT_Conv_S210_Command";
      GC01_FB15 : "UDT_Conv_G115D_Command";
      GC01_FB16 : "UDT_Conv_G115D_Command";
      GC01_FB17 : "UDT_Conv_G115D_Command";
      GC01_FB18 : "UDT_Conv_G115D_Command";
      GC01_FB19 : "UDT_Conv_G115D_Command";
      GC01_FB20 : "UDT_Conv_G115D_Command";
      GC01_FB21 : "UDT_Conv_G115D_Command";
      GC01_FB22 : "UDT_Conv_G115D_Command";
      GC01_FB23 : "UDT_Conv_G115D_Command";
      GC01_FB24 : "UDT_Conv_G115D_Command";
      GC01_FB25 : "UDT_Conv_G115D_Command";
      GC01_FB26 : "UDT_Conv_G115D_Command";
      GC01_FB27 : "UDT_Conv_G115D_Command";
      GC01_FB28 : "UDT_Conv_S210_Command";
      GC01_FB29 : "UDT_Conv_S210_Command";
      GC01_FB30 : "UDT_Conv_S210_Command";
      GC01_FB31 : "UDT_Conv_S210_Command";
      GC01_FB32 : "UDT_Conv_G115D_Command";
      GC02_FB01 : "UDT_Conv_G115D_Command";
      GC02_FB02 : "UDT_Conv_G115D_Command";
      GC02_FB03 : "UDT_Conv_S210_Command";
      GC02_FB04 : "UDT_Conv_S210_Command";
      DT02 : "UDT_Conv_SWS_Command";
      GC02_RC05 : "UDT_Conv_MultiControl_Command";
      GC02_FB06 : "UDT_Conv_G115D_Command";
      GC02_FB07 : "UDT_Conv_G115D_Command";
      GC02_FB08 : "UDT_Conv_G115D_Command";
      GC02_FB09 : "UDT_Conv_G115D_Command";
      GC02_FB10 : "UDT_Conv_G115D_Command";
      GC02_FB11 : "UDT_Conv_G115D_Command";
      GC02_FB12 : "UDT_Conv_G115D_Command";
      GC02_FB13 : "UDT_Conv_G115D_Command";
      GC02_FB14 : "UDT_Conv_G115D_Command";
      GC02_SK15 : "UDT_Conv_G115D_Command";
      GC02_FB16 : "UDT_Conv_S210_Command";
      GC02_FB17 : "UDT_Conv_S210_Command";
      GC02_FB18 : "UDT_Conv_S210_Command";
      GC03_RC01 : "UDT_Conv_MultiControl_Command";
      GC03_RC40 : "UDT_Conv_MultiControl_Command";
      GC03_RC02 : "UDT_Conv_MultiControl_Command";
      GC03_RC03 : "UDT_Conv_MultiControl_Command";
      GC03_RC41 : "UDT_Conv_MultiControl_Command";
      GC03_RC04 : "UDT_Conv_MultiControl_Command";
      GC03_HB05_Merge : "UDT_Merge_2_To_1_Command";
      GC03_HB05 : "UDT_Conv_G115D_Command";
      GC03_FB06 : "UDT_Conv_G115D_Command";
      GC03_FB42 : "UDT_Conv_G115D_Command";
      GC03_FB07 : "UDT_Conv_G115D_Command";
      GC03_FB08 : "UDT_Conv_G115D_Command";
      GC03_FB09 : "UDT_Conv_G115D_Command";
      GC03_FB10 : "UDT_Conv_S210_Command";
      GC03_FB11 : "UDT_Conv_S210_Command";
      DT03 : "UDT_Conv_SWS_Command";
      GC03_RC12 : "UDT_Conv_MultiControl_Command";
      GC03_FB13 : "UDT_Conv_G115D_Command";
      GC03_FB14 : "UDT_Conv_S210_Command";
      GC03_FB15 : "UDT_Conv_S210_Command";
      GC03_FB16 : "UDT_Conv_S210_Command";
      GC03_FB17 : "UDT_Conv_S210_Command";
      GC03_FB18 : "UDT_Conv_G115D_Command";
      GC03_RC19 : "UDT_Conv_G115D_Command";
      GC03_RC20 : "UDT_Conv_MultiControl_Command";
      GC03_FB21_Accmulation : "UDT_Accmulation_Command";
      GC03_FB21 : "UDT_Conv_G115D_Command";
      GC03_FB22 : "UDT_Conv_G115D_Command";
      GC03_FB23 : "UDT_Conv_G115D_Command";
      GC03_FB24 : "UDT_Conv_G115D_Command";
      GC03_FB25 : "UDT_Conv_G115D_Command";
      GC03_FB26 : "UDT_Conv_G115D_Command";
      GC03_FB27 : "UDT_Conv_G115D_Command";
      GC03_FB28 : "UDT_Conv_G115D_Command";
      GC03_FB29 : "UDT_Conv_G115D_Command";
      GC03_FB30 : "UDT_Conv_G115D_Command";
      GC03_FB31 : "UDT_Conv_G115D_Command";
      GC03_FB32_Infeed : "UDT_Induct_On_Gap_Command";
      GC03_FB32 : "UDT_Conv_G115D_Command";
      GC03_RC33 : "UDT_Conv_Dual_G115D_Command";
      GC04_FB04 : "UDT_Conv_G115D_Command";
      GC04_FB05 : "UDT_Conv_G115D_Command";
      GC04_FB06 : "UDT_Conv_G115D_Command";
      GC04_FB07 : "UDT_Conv_G115D_Command";
      GC04_FB08 : "UDT_Conv_G115D_Command";
      GC04_FB09 : "UDT_Conv_G115D_Command";
      GC04_FB10 : "UDT_Conv_S210_Command";
      GC04_FB11 : "UDT_Conv_S210_Command";
      DT04 : "UDT_Conv_SWS_Command";
      GC04_FB12 : "UDT_Conv_G115D_Command";
      GC04_FB13 : "UDT_Conv_G115D_Command";
      GC04_FB14 : "UDT_Conv_G115D_Command";
      GC04_FB15 : "UDT_Conv_G115D_Command";
      GC04_FB16 : "UDT_Conv_G115D_Command";
      GC04_FB17 : "UDT_Conv_G115D_Command";
      GC04_FB18 : "UDT_Conv_G115D_Command";
      GC04_FB19 : "UDT_Conv_G115D_Command";
      GC04_RC20 : "UDT_Conv_MultiControl_Command";
      GC04_RC21 : "UDT_Conv_Dual_G115D_Command";
      GC05_RC01 : "UDT_Conv_MultiControl_Command";
      GC05_RC02 : "UDT_Conv_MultiControl_Command";
      GC05_RC03 : "UDT_Conv_MultiControl_Command";
      GC05_RC10 : "UDT_Conv_MultiControl_Command";
      GC05_FB04 : "UDT_Conv_G115D_Command";
      GC05_FB05 : "UDT_Conv_G115D_Command";
      GC05_RC06 : "UDT_Conv_MultiControl_Command";
      GC05_RC07 : "UDT_Conv_G115D_Command";
      GC06_RC01 : "UDT_Conv_MultiControl_Command";
      GC06_FB02 : "UDT_Conv_G115D_Command";
      GC06_FB03 : "UDT_Conv_G115D_Command";
      GC06_RC04_Merge : "UDT_Merge_3_To_1_Command";
      GC06_RC04 : "UDT_Conv_Triple_G115D_Command";
      GC06_FB05 : "UDT_Conv_G115D_Command";
      GC06_FB06 : "UDT_Conv_G115D_Command";
      GC06_FB07 : "UDT_Conv_G115D_Command";
      GC06_SK08 : "UDT_Conv_G115D_Command";
      GC07_FB01 : "UDT_Conv_G115D_Command";
      GC07_RC02 : "UDT_Conv_Dual_G115D_Command";
      GC07_RC03 : "UDT_Conv_MultiControl_Command";
      GC07_RC04 : "UDT_Conv_MultiControl_Command";
      GC07_RC05 : "UDT_Conv_MultiControl_Command";
      GC07_RC06 : "UDT_Conv_MultiControl_Command";
      GC07_RC10 : "UDT_Conv_MultiControl_Command";
      GC07_RC07 : "UDT_Conv_MultiControl_Command";
      GC07_RC08 : "UDT_Conv_MultiControl_Command";
      GC07_RC11 : "UDT_Conv_MultiControl_Command";
      GC07_FB09 : "UDT_Conv_G115D_Command";
   END_STRUCT;


BEGIN

END_DATA_BLOCK

DATA_BLOCK "DI_GC02_FB16_Conv_S210"
{ S7_Optimized_Access := 'TRUE' }
VERSION : 0.1
NON_RETAIN
"FB_Conv_S210"

BEGIN

END_DATA_BLOCK

FUNCTION "FC_Inbound_Line2" : Void
{ S7_Optimized_Access := 'TRUE' }
VERSION : 0.1
   VAR_TEMP
      t_SWS_Trigger : Bool;
      t_Fnd_Items : Int;
      t_Fnd_Entry : Int;
      t_Fnd_Data : Int;
      t_Int_Not_Used : Int;
   END_VAR


BEGIN
	REGION NETWORK: GC02_FB01 - Transport Conveyor - G115D

	    // FB_Conv_G115D
	    "DI_GC02_FB01_Conv_G115D"(i_Telegram_HW_ID   := "=MHE+GC02_FB01~PROFINET_interface~Standard_telegram_1",
	                              i_Additional_HW_ID := "=MHE+GC02_FB01~PROFINET_interface~Annex_Free_telegram",
	                              i_IO_PEC_Position  := TRUE,
	                              i_IO_PEC_Trigger   := TRUE,
	                              i_Setting          := "DB_Setting".GC02_FB01,
	                              i_External_Request := "DB_External".GC02_FB01,
	                              i_Command          := "DB_Command".GC02_FB01,
	                              o_Status           => "DB_Status".GC02_FB01,
	                              o_General_Status   => "DB_General_Status".GC02_FB01,
	                              o_Diagnostics      => "DB_Diagnostics".GC02_FB01,
	                              io_Global          := "DB_Global",
	                              io_System_Control  := "DB_System_Control".GC02_FB01,
	                              io_G115D_IO        := "DB_IO".GC02_FB01,
	                              io_FIF_Upstream    := "DB_Flow_Interface".Upstream_Dummy,
	                              io_FIF             := "DB_Flow_Interface".GC02_FB01,
	                              io_FIF_Downstream  := "DB_Flow_Interface".GC02_FB02);

	END_REGION

	REGION NETWORK: GC02_FB02 - Transport Conveyor - G115D

	    // FB_Conv_G115D
	    "DI_GC02_FB02_Conv_G115D"(i_Telegram_HW_ID   := "=MHE+GC02_FB02~PROFINET_interface~Standard_telegram_1",
	                              i_Additional_HW_ID := "=MHE+GC02_FB02~PROFINET_interface~Annex_Free_telegram",
	                              i_IO_PEC_Position  := TRUE,
	                              i_IO_PEC_Trigger   := TRUE,
	                              i_Setting          := "DB_Setting".GC02_FB02,
	                              i_External_Request := "DB_External".GC02_FB02,
	                              i_Command          := "DB_Command".GC02_FB02,
	                              o_Status           => "DB_Status".GC02_FB02,
	                              o_General_Status   => "DB_General_Status".GC02_FB02,
	                              o_Diagnostics      => "DB_Diagnostics".GC02_FB02,
	                              io_Global          := "DB_Global",
	                              io_System_Control  := "DB_System_Control".GC02_FB02,
	                              io_G115D_IO        := "DB_IO".GC02_FB02,
	                              io_FIF_Upstream    := "DB_Flow_Interface".GC02_FB01,
	                              io_FIF             := "DB_Flow_Interface".GC02_FB02,
	                              io_FIF_Downstream  := "DB_Flow_Interface".Downstream_Dummy);

	END_REGION

	REGION NETWORK: GC02_FB03 - Transport Conveyor - S210

	    // FB_Conv_S210
	    "DI_GC02_FB03_Conv_S210"(i_Telegram_HW_ID   := "=MHE+GC02_FB03~PROFINET_interface~Drive_control_SIEMENS_teleg,,,",
	                             i_Additional_HW_ID := "=MHE+GC02_FB03~PROFINET_interface~Drive_control_Annex_Free_te,,,",
	                             i_IO_PEC_Position  := TRUE,
	                             i_IO_PEC_Trigger   := TRUE,
	                             i_Setting          := "DB_Setting".GC02_FB03,
	                             i_Command          := "DB_Command".GC02_FB03,
	                             i_External_Request := "DB_External".GC02_FB03,
	                             o_Status           => "DB_Status".GC02_FB03,
	                             o_General_Status   => "DB_General_Status".GC02_FB03,
	                             o_Diagnostics      => "DB_Diagnostics".GC02_FB03,
	                             io_Global          := "DB_Global",
	                             io_System_Control  := "DB_System_Control".GC02_FB03,
	                             io_S210_IO         := "DB_IO".GC02_FB03,
	                             io_FIF_Upstream    := "DB_Flow_Interface".Upstream_Dummy,
	                             io_FIF             := "DB_Flow_Interface".GC02_FB03,
	                             io_FIF_Downstream  := "DB_Flow_Interface".GC02_FB04);

	END_REGION

	REGION NETWORK: GC02_FB04 - Transport Conveyor - S210

	    // FB_Conv_S210
	    "DI_GC02_FB04_Conv_S210"(i_Telegram_HW_ID   := "=MHE+GC02_FB04~PROFINET_interface~Drive_control_SIEMENS_teleg,,,",
	                             i_Additional_HW_ID := "=MHE+GC02_FB04~PROFINET_interface~Drive_control_Annex_Free_te,,,",
	                             i_IO_PEC_Position  := TRUE,
	                             i_IO_PEC_Trigger   := TRUE,
	                             i_Setting          := "DB_Setting".GC02_FB04,
	                             i_Command          := "DB_Command".GC02_FB04,
	                             i_External_Request := "DB_External".GC02_FB04,
	                             o_Status           => "DB_Status".GC02_FB04,
	                             o_General_Status   => "DB_General_Status".GC02_FB04,
	                             o_Diagnostics      => "DB_Diagnostics".GC02_FB04,
	                             io_Global          := "DB_Global",
	                             io_System_Control  := "DB_System_Control".GC02_FB04,
	                             io_S210_IO         := "DB_IO".GC02_FB04,
	                             io_FIF_Upstream    := "DB_Flow_Interface".GC02_FB03,
	                             io_FIF             := "DB_Flow_Interface".GC02_FB04,
	                             io_FIF_Downstream  := "DB_Flow_Interface".DT02);

	END_REGION

	REGION NETWORK: DT02 - Steerable Wheel Sorter

	    // FB_Conv_SWS
	    "DI_DT02_Conv_SWS"(i_New_Item_Present            := FALSE,
	                       i_CMD_Divert_Left             := FALSE,
	                       i_CMD_Divert_Straight         := FALSE,
	                       i_CMD_Divert_Right            := FALSE,
	                       i_Setting                     := "DB_Setting".DT02,
	                       i_External_Request            := "DB_External".DT02,
	                       i_U401_Additional_HW_ID       := "=MHE+AC03_U401~PROFINET_Interface~Drive_Control_Annex_Free_te,,,",
	                       i_U401_Telegram_HW_ID         := "=MHE+AC03_U401~PROFINET_Interface~Drive_Control_SIEMENS_teleg,,,",
	                       i_U411_Additional_HW_ID       := "=MHE+AC03_U411~PROFINET_Interface~Drive_Control_Annex_Free_te,,,",
	                       i_U411_Telegram_HW_ID         := "=MHE+AC03_U411~PROFINET_Interface~Drive_Control_SIEMENS_teleg,,,",
	                       i_U421_Additional_HW_ID       := "=MHE+AC03_U421~PROFINET_Interface~Drive_Control_Annex_Free_te,,,",
	                       i_U421_Telegram_HW_ID         := "=MHE+AC03_U421~PROFINET_Interface~Drive_Control_SIEMENS_teleg,,,",
	                       i_U431_Additional_HW_ID       := "=MHE+AC03_U431~PROFINET_Interface~Drive_Control_Annex_Free_te,,,",
	                       i_U431_Telegram_HW_ID         := "=MHE+AC03_U431~PROFINET_Interface~Drive_Control_SIEMENS_teleg,,,",
	                       i_U441_Additional_HW_ID       := "=MHE+AC03_U441~PROFINET_Interface~Drive_Control_Annex_Free_te,,,",
	                       i_U441_Telegram_HW_ID         := "=MHE+AC03_U441~PROFINET_Interface~Drive_Control_SIEMENS_teleg,,,",
	                       i_U451_Additional_HW_ID       := "=MHE+AC03_U451~PROFINET_Interface~Drive_Control_Annex_Free_te,,,",
	                       i_U451_Telegram_HW_ID         := "=MHE+AC03_U451~PROFINET_Interface~Drive_Control_SIEMENS_teleg,,,",
	                       i_U461_Additional_HW_ID       := "=MHE+AC03_U461~PROFINET_Interface~Drive_Control_Annex_Free_te,,,",
	                       i_U461_Telegram_HW_ID         := "=MHE+AC03_U461~PROFINET_Interface~Drive_Control_SIEMENS_teleg,,,",
	                       i_U471_Additional_HW_ID       := "=MHE+AC03_U471~PROFINET_Interface~Drive_Control_Annex_Free_te,,,",
	                       i_U471_Telegram_HW_ID         := "=MHE+AC03_U471~PROFINET_Interface~Drive_Control_SIEMENS_teleg,,,",
	                       i_U481_Additional_HW_ID       := "=MHE+AC03_U481~PROFINET_Interface~Drive_Control_Annex_Free_te,,,",
	                       i_U481_Telegram_HW_ID         := "=MHE+AC03_U481~PROFINET_Interface~Drive_Control_SIEMENS_teleg,,,",
	                       i_Roller_Gateway_Input_HW_ID  := "=MHE+AC03_NT100~Input",
	                       i_Roller_Gateway_Output_HW_ID := "=MHE+AC03_NT100~Output",
	                       o_Status                      => "DB_Status".DT02,
	                       o_General_Status              => "DB_General_Status".DT02,
	                       io_Global                     := "DB_Global",
	                       io_System_Control             := "DB_System_Control".DT02,
	                       io_Interface                  := "DB_IO".DT02,
	                       io_Gateway_Interface          := "DB_IO".AC03_NT100,
	                       io_Command                    := "DB_Command".DT02,
	                       io_FIF_Upstream               := "DB_Flow_Interface".GC02_FB04,
	                       io_FIF                        := "DB_Flow_Interface".DT02,
	                       io_FIF_Downstream             := "DB_Flow_Interface".GC02_RC05);

	END_REGION

	REGION NETWORK: GC02_RC05 - Transport Conveyor - Interroll MultiControl

	    // FB_Conv_MultiControl
	    "DI_GC02_RC05_Conv_MultiControl"(i_IO_PEC_Position      := TRUE,
	                                     i_IO_PEC_Trigger       := TRUE,
	                                     i_Setting              := "DB_Setting".GC02_RC05,
	                                     i_External_Request     := "DB_External".GC02_RC05,
	                                     i_Command              := "DB_Command".GC02_RC05,
	                                     o_Status               => "DB_Status".GC02_RC05,
	                                     o_General_Status       => "DB_General_Status".GC02_RC05,
	                                     o_Diagnostics          => "DB_Diagnostics".GC02_RC05,
	                                     io_Global              := "DB_Global",
	                                     io_System_Control      := "DB_System_Control".GC02_RC05,
	                                     io_MultiControl_U01_IO := "DB_IO".GC02_RC05_A01,
	                                     io_MultiControl_U02_IO := "DB_IO".MultiControl_Dummy,
	                                     io_MultiControl_U03_IO := "DB_IO".MultiControl_Dummy,
	                                     io_MultiControl_U04_IO := "DB_IO".MultiControl_Dummy,
	                                     io_FIF_Upstream        := "DB_Flow_Interface".DT02,
	                                     io_FIF                 := "DB_Flow_Interface".GC02_RC05,
	                                     io_FIF_Downstream      := "DB_Flow_Interface".GC02_FB06);

	END_REGION

	REGION NETWORK: GC02_FB06 - Transport Conveyor - G115D

	    // FB_Conv_G115D
	    "DI_GC02_FB06_Conv_G115D"(i_Telegram_HW_ID   := "=MHE+GC02_FB06~PROFINET_interface~Standard_telegram_1",
	                              i_Additional_HW_ID := "=MHE+GC02_FB06~PROFINET_interface~Annex_Free_telegram",
	                              i_IO_PEC_Position  := TRUE,
	                              i_IO_PEC_Trigger   := TRUE,
	                              i_Setting          := "DB_Setting".GC02_FB06,
	                              i_External_Request := "DB_External".GC02_FB06,
	                              i_Command          := "DB_Command".GC02_FB06,
	                              o_Status           => "DB_Status".GC02_FB06,
	                              o_General_Status   => "DB_General_Status".GC02_FB06,
	                              o_Diagnostics      => "DB_Diagnostics".GC02_FB06,
	                              io_Global          := "DB_Global",
	                              io_System_Control  := "DB_System_Control".GC02_FB06,
	                              io_G115D_IO        := "DB_IO".GC02_FB06,
	                              io_FIF_Upstream    := "DB_Flow_Interface".GC02_RC05,
	                              io_FIF             := "DB_Flow_Interface".GC02_FB06,
	                              io_FIF_Downstream  := "DB_Flow_Interface".GC02_FB07);

	END_REGION

	REGION NETWORK: GC02_FB07 - Transport Conveyor - G115D

	    // FB_Conv_G115D
	    "DI_GC02_FB07_Conv_G115D"(i_Telegram_HW_ID   := "=MHE+GC02_FB07~PROFINET_interface~Standard_telegram_1",
	                              i_Additional_HW_ID := "=MHE+GC02_FB07~PROFINET_interface~Annex_Free_telegram",
	                              i_IO_PEC_Position  := TRUE,
	                              i_IO_PEC_Trigger   := TRUE,
	                              i_Setting          := "DB_Setting".GC02_FB07,
	                              i_External_Request := "DB_External".GC02_FB07,
	                              i_Command          := "DB_Command".GC02_FB07,
	                              o_Status           => "DB_Status".GC02_FB07,
	                              o_General_Status   => "DB_General_Status".GC02_FB07,
	                              o_Diagnostics      => "DB_Diagnostics".GC02_FB07,
	                              io_Global          := "DB_Global",
	                              io_System_Control  := "DB_System_Control".GC02_FB07,
	                              io_G115D_IO        := "DB_IO".GC02_FB07,
	                              io_FIF_Upstream    := "DB_Flow_Interface".GC02_FB06,
	                              io_FIF             := "DB_Flow_Interface".GC02_FB07,
	                              io_FIF_Downstream  := "DB_Flow_Interface".GC02_FB08);

	END_REGION

	REGION NETWORK: GC02_FB08 - Transport Conveyor - G115D

	    // FB_Conv_G115D
	    "DI_GC02_FB08_Conv_G115D"(i_Telegram_HW_ID   := "=MHE+GC02_FB08~PROFINET_interface~Standard_telegram_1",
	                              i_Additional_HW_ID := "=MHE+GC02_FB08~PROFINET_interface~Annex_Free_telegram",
	                              i_IO_PEC_Position  := TRUE,
	                              i_IO_PEC_Trigger   := TRUE,
	                              i_Setting          := "DB_Setting".GC02_FB08,
	                              i_External_Request := "DB_External".GC02_FB08,
	                              i_Command          := "DB_Command".GC02_FB08,
	                              o_Status           => "DB_Status".GC02_FB08,
	                              o_General_Status   => "DB_General_Status".GC02_FB08,
	                              o_Diagnostics      => "DB_Diagnostics".GC02_FB08,
	                              io_Global          := "DB_Global",
	                              io_System_Control  := "DB_System_Control".GC02_FB08,
	                              io_G115D_IO        := "DB_IO".GC02_FB08,
	                              io_FIF_Upstream    := "DB_Flow_Interface".GC02_FB07,
	                              io_FIF             := "DB_Flow_Interface".GC02_FB08,
	                              io_FIF_Downstream  := "DB_Flow_Interface".GC04_RC21);

	END_REGION

	REGION NETWORK: GC04_RC21 - Transport Conveyor - Dual G115D

	    // FB_Conv_Dual_G115D
	    "DI_GC04_RC21_Conv_Dual_G115D"(i_U01_Telegram_HW_ID   := "=MHE+GC04_RC21_M01~PROFINET_interface~Standard_telegram_1",
	                                   i_U01_Additional_HW_ID := "=MHE+GC04_RC21_M01~PROFINET_interface~Annex_Free_telegram",
	                                   i_U02_Telegram_HW_ID   := "=MHE+GC04_RC21_M02~PROFINET_interface~Standard_telegram_1",
	                                   i_U02_Additional_HW_ID := "=MHE+GC04_RC21_M02~PROFINET_interface~Annex_Free_telegram",
	                                   i_IO_PEC_Position      := TRUE,
	                                   i_IO_PEC_Trigger       := TRUE,
	                                   i_Setting              := "DB_Setting".GC04_RC21,
	                                   i_External_Request     := "DB_External".GC04_RC21,
	                                   i_Command              := "DB_Command".GC04_RC21,
	                                   o_Status               => "DB_Status".GC04_RC21,
	                                   o_General_Status       => "DB_General_Status".GC04_RC21,
	                                   o_Diagnostics          => "DB_Diagnostics".GC04_RC21,
	                                   io_Global              := "DB_Global",
	                                   io_System_Control      := "DB_System_Control".GC04_RC21,
	                                   io_U01_G115D_IO        := "DB_IO".GC04_RC21_M01,
	                                   io_U02_G115D_IO        := "DB_IO".GC04_RC21_M02,
	                                   io_FIF_Upstream        := "DB_Flow_Interface".GC02_FB08,
	                                   io_FIF                 := "DB_Flow_Interface".GC04_RC21,
	                                   io_FIF_Downstream      := "DB_Flow_Interface".GC02_FB09);

	END_REGION

	REGION NETWORK: GC02_FB09 - Transport Conveyor - G115D

	    // FB_Conv_G115D
	    "DI_GC02_FB09_Conv_G115D"(i_Telegram_HW_ID   := "=MHE+GC02_FB09~PROFINET_interface~Standard_telegram_1",
	                              i_Additional_HW_ID := "=MHE+GC02_FB09~PROFINET_interface~Annex_Free_telegram",
	                              i_IO_PEC_Position  := TRUE,
	                              i_IO_PEC_Trigger   := TRUE,
	                              i_Setting          := "DB_Setting".GC02_FB09,
	                              i_External_Request := "DB_External".GC02_FB09,
	                              i_Command          := "DB_Command".GC02_FB09,
	                              o_Status           => "DB_Status".GC02_FB09,
	                              o_General_Status   => "DB_General_Status".GC02_FB09,
	                              o_Diagnostics      => "DB_Diagnostics".GC02_FB09,
	                              io_Global          := "DB_Global",
	                              io_System_Control  := "DB_System_Control".GC02_FB09,
	                              io_G115D_IO        := "DB_IO".GC02_FB09,
	                              io_FIF_Upstream    := "DB_Flow_Interface".GC04_RC21,
	                              io_FIF             := "DB_Flow_Interface".GC02_FB09,
	                              io_FIF_Downstream  := "DB_Flow_Interface".GC02_FB10);

	END_REGION

	REGION NETWORK: GC02_FB10 - Transport Conveyor - G115D

	    // FB_Conv_G115D
	    "DI_GC02_FB10_Conv_G115D"(i_Telegram_HW_ID   := "=MHE+GC02_FB10~PROFINET_interface~Standard_telegram_1",
	                              i_Additional_HW_ID := "=MHE+GC02_FB10~PROFINET_interface~Annex_Free_telegram",
	                              i_IO_PEC_Position  := TRUE,
	                              i_IO_PEC_Trigger   := TRUE,
	                              i_Setting          := "DB_Setting".GC02_FB10,
	                              i_External_Request := "DB_External".GC02_FB10,
	                              i_Command          := "DB_Command".GC02_FB10,
	                              o_Status           => "DB_Status".GC02_FB10,
	                              o_General_Status   => "DB_General_Status".GC02_FB10,
	                              o_Diagnostics      => "DB_Diagnostics".GC02_FB10,
	                              io_Global          := "DB_Global",
	                              io_System_Control  := "DB_System_Control".GC02_FB10,
	                              io_G115D_IO        := "DB_IO".GC02_FB10,
	                              io_FIF_Upstream    := "DB_Flow_Interface".GC02_FB09,
	                              io_FIF             := "DB_Flow_Interface".GC02_FB10,
	                              io_FIF_Downstream  := "DB_Flow_Interface".GC02_FB11);

	END_REGION

	REGION NETWORK: GC02_FB11 - Transport Conveyor - G115D

	    // FB_Conv_G115D
	    "DI_GC02_FB11_Conv_G115D"(i_Telegram_HW_ID   := "=MHE+GC02_FB11~PROFINET_interface~Standard_telegram_1",
	                              i_Additional_HW_ID := "=MHE+GC02_FB11~PROFINET_interface~Annex_Free_telegram",
	                              i_IO_PEC_Position  := TRUE,
	                              i_IO_PEC_Trigger   := TRUE,
	                              i_Setting          := "DB_Setting".GC02_FB11,
	                              i_External_Request := "DB_External".GC02_FB11,
	                              i_Command          := "DB_Command".GC02_FB11,
	                              o_Status           => "DB_Status".GC02_FB11,
	                              o_General_Status   => "DB_General_Status".GC02_FB11,
	                              o_Diagnostics      => "DB_Diagnostics".GC02_FB11,
	                              io_Global          := "DB_Global",
	                              io_System_Control  := "DB_System_Control".GC02_FB11,
	                              io_G115D_IO        := "DB_IO".GC02_FB11,
	                              io_FIF_Upstream    := "DB_Flow_Interface".GC02_FB10,
	                              io_FIF             := "DB_Flow_Interface".GC02_FB11,
	                              io_FIF_Downstream  := "DB_Flow_Interface".GC02_FB12);

	END_REGION

	REGION NETWORK: GC02_FB12 - Transport Conveyor - G115D

	    // FB_Conv_G115D
	    "DI_GC02_FB12_Conv_G115D"(i_Telegram_HW_ID   := "=MHE+GC02_FB12~PROFINET_interface~Standard_telegram_1",
	                              i_Additional_HW_ID := "=MHE+GC02_FB12~PROFINET_interface~Annex_Free_telegram",
	                              i_IO_PEC_Position  := TRUE,
	                              i_IO_PEC_Trigger   := TRUE,
	                              i_Setting          := "DB_Setting".GC02_FB12,
	                              i_External_Request := "DB_External".GC02_FB12,
	                              i_Command          := "DB_Command".GC02_FB12,
	                              o_Status           => "DB_Status".GC02_FB12,
	                              o_General_Status   => "DB_General_Status".GC02_FB12,
	                              o_Diagnostics      => "DB_Diagnostics".GC02_FB12,
	                              io_Global          := "DB_Global",
	                              io_System_Control  := "DB_System_Control".GC02_FB12,
	                              io_G115D_IO        := "DB_IO".GC02_FB12,
	                              io_FIF_Upstream    := "DB_Flow_Interface".GC02_FB11,
	                              io_FIF             := "DB_Flow_Interface".GC02_FB12,
	                              io_FIF_Downstream  := "DB_Flow_Interface".GC02_FB13);

	END_REGION

	REGION NETWORK: GC02_FB13 - Transport Conveyor - G115D

	    // FB_Conv_G115D
	    "DI_GC02_FB13_Conv_G115D"(i_Telegram_HW_ID   := "=MHE+GC02_FB13~PROFINET_interface~Standard_telegram_1",
	                              i_Additional_HW_ID := "=MHE+GC02_FB13~PROFINET_interface~Annex_Free_telegram",
	                              i_IO_PEC_Position  := TRUE,
	                              i_IO_PEC_Trigger   := TRUE,
	                              i_Setting          := "DB_Setting".GC02_FB13,
	                              i_External_Request := "DB_External".GC02_FB13,
	                              i_Command          := "DB_Command".GC02_FB13,
	                              o_Status           => "DB_Status".GC02_FB13,
	                              o_General_Status   => "DB_General_Status".GC02_FB13,
	                              o_Diagnostics      => "DB_Diagnostics".GC02_FB13,
	                              io_Global          := "DB_Global",
	                              io_System_Control  := "DB_System_Control".GC02_FB13,
	                              io_G115D_IO        := "DB_IO".GC02_FB13,
	                              io_FIF_Upstream    := "DB_Flow_Interface".GC02_FB12,
	                              io_FIF             := "DB_Flow_Interface".GC02_FB13,
	                              io_FIF_Downstream  := "DB_Flow_Interface".GC02_FB14);

	END_REGION

	REGION NETWORK: GC02_FB14 - Transport Conveyor - G115D

	    // FB_Conv_G115D
	    "DI_GC02_FB14_Conv_G115D"(i_Telegram_HW_ID   := "=MHE+GC02_FB14~PROFINET_interface~Standard_telegram_1",
	                              i_Additional_HW_ID := "=MHE+GC02_FB14~PROFINET_interface~Annex_Free_telegram",
	                              i_IO_PEC_Position  := TRUE,
	                              i_IO_PEC_Trigger   := TRUE,
	                              i_Setting          := "DB_Setting".GC02_FB14,
	                              i_External_Request := "DB_External".GC02_FB14,
	                              i_Command          := "DB_Command".GC02_FB14,
	                              o_Status           => "DB_Status".GC02_FB14,
	                              o_General_Status   => "DB_General_Status".GC02_FB14,
	                              o_Diagnostics      => "DB_Diagnostics".GC02_FB14,
	                              io_Global          := "DB_Global",
	                              io_System_Control  := "DB_System_Control".GC02_FB14,
	                              io_G115D_IO        := "DB_IO".GC02_FB14,
	                              io_FIF_Upstream    := "DB_Flow_Interface".GC02_FB13,
	                              io_FIF             := "DB_Flow_Interface".GC02_FB14,
	                              io_FIF_Downstream  := "DB_Flow_Interface".GC02_SK15);

	END_REGION

	REGION NETWORK: GC02_SK15 - Transport Conveyor - G115D

	    // FB_Conv_G115D
	    "DI_GC02_SK15_Conv_G115D"(i_Telegram_HW_ID   := "=MHE+GC02_SK15~PROFINET_interface~Standard_telegram_1",
	                              i_Additional_HW_ID := "=MHE+GC02_SK15~PROFINET_interface~Annex_Free_telegram",
	                              i_IO_PEC_Position  := TRUE,
	                              i_IO_PEC_Trigger   := TRUE,
	                              i_Setting          := "DB_Setting".GC02_SK15,
	                              i_External_Request := "DB_External".GC02_SK15,
	                              i_Command          := "DB_Command".GC02_SK15,
	                              o_Status           => "DB_Status".GC02_SK15,
	                              o_General_Status   => "DB_General_Status".GC02_SK15,
	                              o_Diagnostics      => "DB_Diagnostics".GC02_SK15,
	                              io_Global          := "DB_Global",
	                              io_System_Control  := "DB_System_Control".GC02_SK15,
	                              io_G115D_IO        := "DB_IO".GC02_SK15,
	                              io_FIF_Upstream    := "DB_Flow_Interface".GC02_FB14,
	                              io_FIF             := "DB_Flow_Interface".GC02_SK15,
	                              io_FIF_Downstream  := "DB_Flow_Interface".GC02_FB16);

	END_REGION

	REGION NETWORK: GC02_FB16 - Transport Conveyor - S210

	    // FB_Conv_S210
	    "DI_GC02_FB16_Conv_S210"(i_Telegram_HW_ID   := "=MHE+GC02_FB16~PROFINET_interface~Drive_control_SIEMENS_teleg,,,",
	                             i_Additional_HW_ID := "=MHE+GC02_FB16~PROFINET_interface~Drive_control_Annex_Free_te,,,",
	                             i_IO_PEC_Position  := TRUE,
	                             i_IO_PEC_Trigger   := TRUE,
	                             i_Setting          := "DB_Setting".GC02_FB16,
	                             i_Command          := "DB_Command".GC02_FB16,
	                             i_External_Request := "DB_External".GC02_FB16,
	                             o_Status           => "DB_Status".GC02_FB16,
	                             o_General_Status   => "DB_General_Status".GC02_FB16,
	                             o_Diagnostics      => "DB_Diagnostics".GC02_FB16,
	                             io_Global          := "DB_Global",
	                             io_System_Control  := "DB_System_Control".GC02_FB16,
	                             io_S210_IO         := "DB_IO".GC02_FB16,
	                             io_FIF_Upstream    := "DB_Flow_Interface".GC02_SK15,
	                             io_FIF             := "DB_Flow_Interface".GC02_FB16,
	                             io_FIF_Downstream  := "DB_Flow_Interface".GC02_FB17);

	END_REGION

	REGION NETWORK: GC02_FB17 - Transport Conveyor - S210

	    // FB_Conv_S210
	    "DI_GC02_FB17_Conv_S210"(i_Telegram_HW_ID   := "=MHE+GC02_FB17~PROFINET_interface~Drive_control_SIEMENS_teleg,,,",
	                             i_Additional_HW_ID := "=MHE+GC02_FB17~PROFINET_interface~Drive_control_Annex_Free_te,,,",
	                             i_IO_PEC_Position  := TRUE,
	                             i_IO_PEC_Trigger   := TRUE,
	                             i_Setting          := "DB_Setting".GC02_FB17,
	                             i_Command          := "DB_Command".GC02_FB17,
	                             i_External_Request := "DB_External".GC02_FB17,
	                             o_Status           => "DB_Status".GC02_FB17,
	                             o_General_Status   => "DB_General_Status".GC02_FB17,
	                             o_Diagnostics      => "DB_Diagnostics".GC02_FB17,
	                             io_Global          := "DB_Global",
	                             io_System_Control  := "DB_System_Control".GC02_FB17,
	                             io_S210_IO         := "DB_IO".GC02_FB17,
	                             io_FIF_Upstream    := "DB_Flow_Interface".GC02_FB16,
	                             io_FIF             := "DB_Flow_Interface".GC02_FB17,
	                             io_FIF_Downstream  := "DB_Flow_Interface".GC02_FB18);

	END_REGION

	REGION NETWORK: GC02_FB18 - Transport Conveyor - S210

	    // FB_Conv_S210
	    "DI_GC02_FB18_Conv_S210"(i_Telegram_HW_ID   := "=MHE+GC02_FB18~PROFINET_interface~Drive_control_SIEMENS_teleg,,,",
	                             i_Additional_HW_ID := "=MHE+GC02_FB18~PROFINET_interface~Drive_control_Annex_Free_te,,,",
	                             i_IO_PEC_Position  := TRUE,
	                             i_IO_PEC_Trigger   := TRUE,
	                             i_Setting          := "DB_Setting".GC02_FB18,
	                             i_Command          := "DB_Command".GC02_FB18,
	                             i_External_Request := "DB_External".GC02_FB18,
	                             o_Status           => "DB_Status".GC02_FB18,
	                             o_General_Status   => "DB_General_Status".GC02_FB18,
	                             o_Diagnostics      => "DB_Diagnostics".GC02_FB18,
	                             io_Global          := "DB_Global",
	                             io_System_Control  := "DB_System_Control".GC02_FB18,
	                             io_S210_IO         := "DB_IO".GC02_FB18,
	                             io_FIF_Upstream    := "DB_Flow_Interface".GC02_FB17,
	                             io_FIF             := "DB_Flow_Interface".GC02_FB18,
	                             io_FIF_Downstream  := "DB_Flow_Interface".Downstream_Dummy);

	END_REGION
END_FUNCTION

